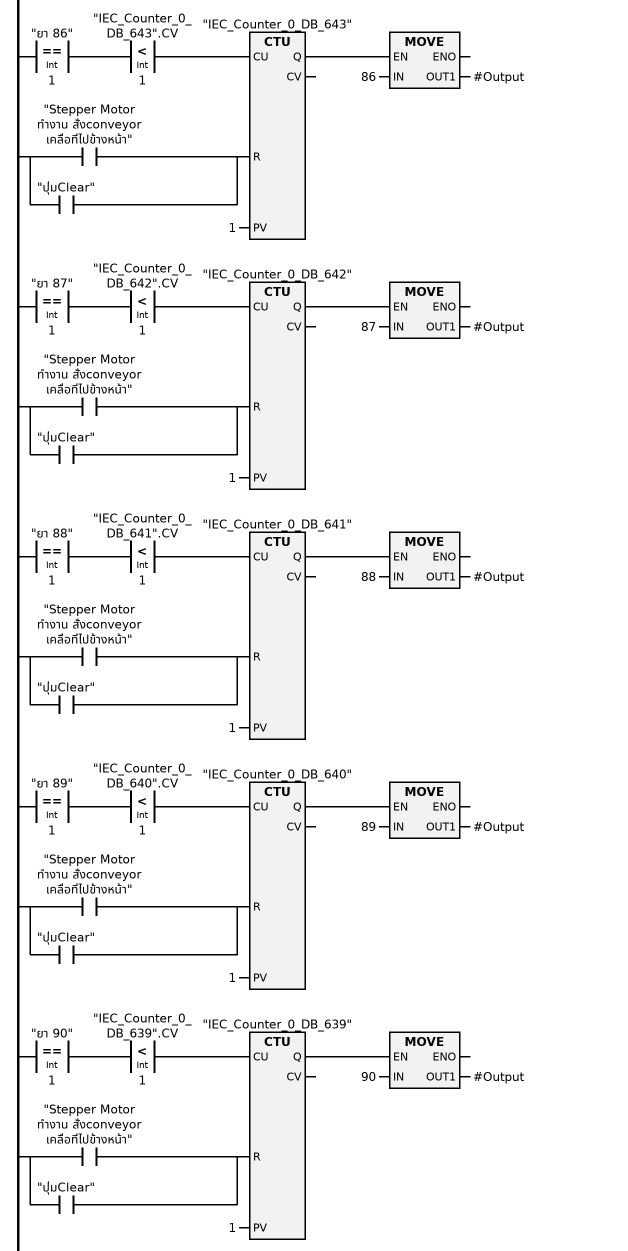
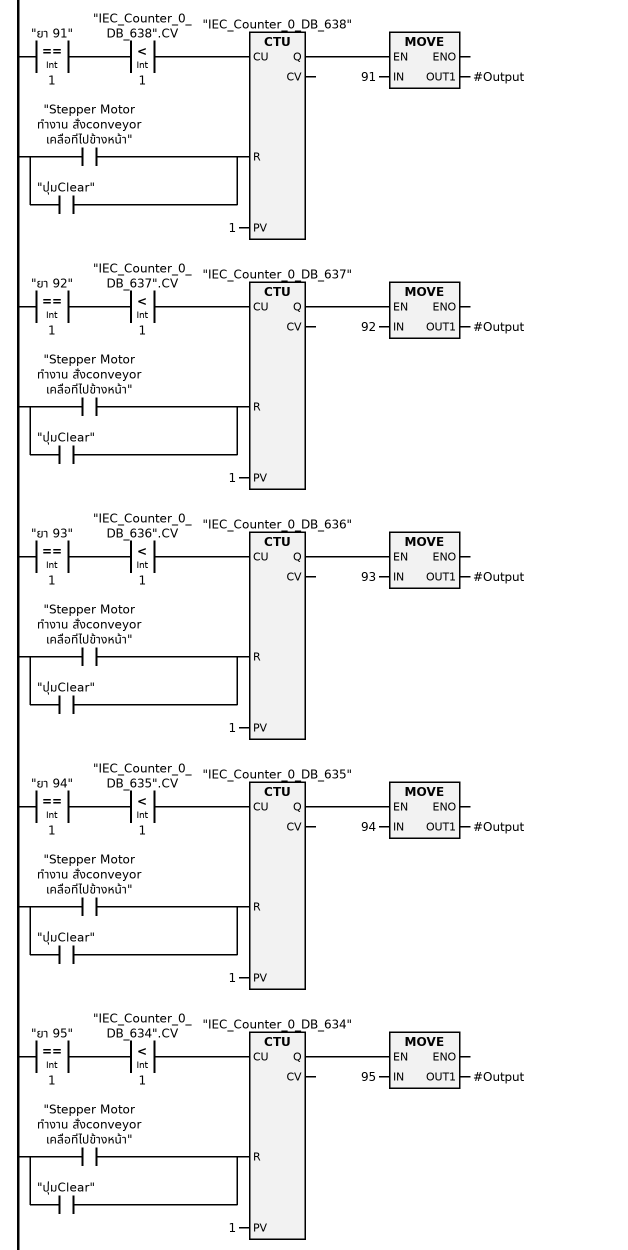
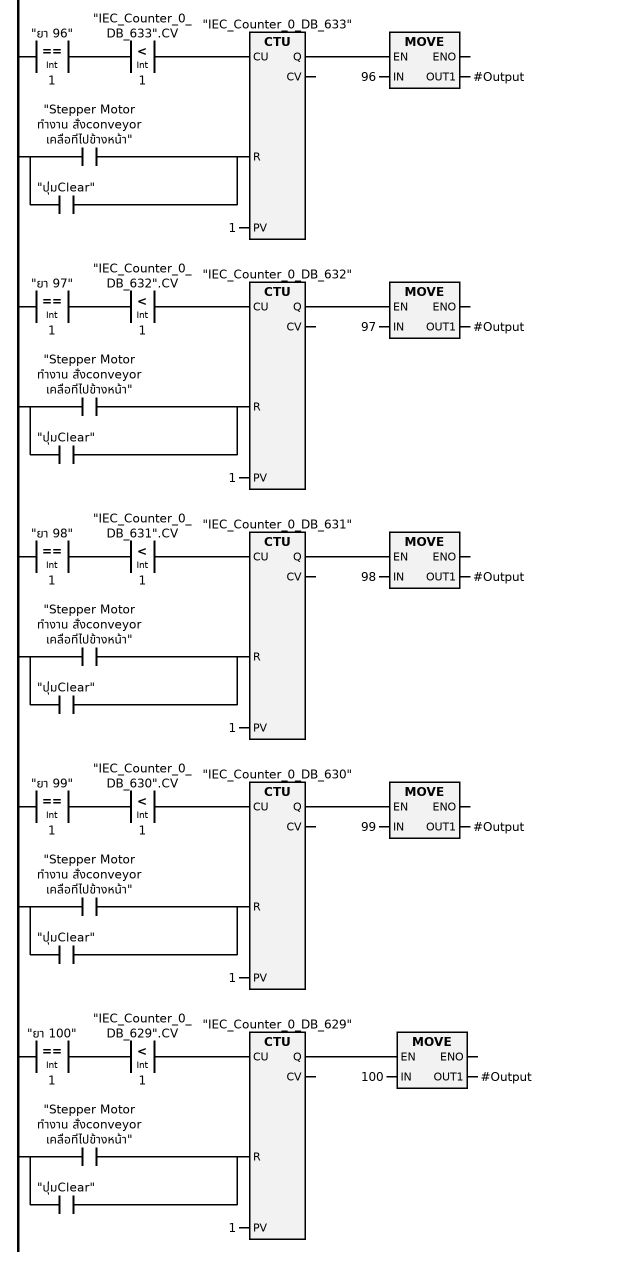
   "IEC_Counter_0_DB_644".CTU(CU := ("ยา 81" = 1) AND ("IEC_Counter_0_DB_644".CV < 1),
                           R := "Stepper Motor ทำงาน สั่งconveyor เคลื่อที่ไปข้างหน้า" OR "ปุ่มClear",
                           PV := 1);
   IF "IEC_Counter_0_DB_644".Q THEN #Output := 81; END_IF;
   "IEC_Counter_0_DB_645".CTU(CU := ("ยา 82" = 1) AND ("IEC_Counter_0_DB_645".CV < 1),
                           R := "Stepper Motor ทำงาน สั่งconveyor เคลื่อที่ไปข้างหน้า" OR "ปุ่มClear",
                           PV := 1);
   IF "IEC_Counter_0_DB_645".Q THEN #Output := 82; END_IF;
   "IEC_Counter_0_DB_647".CTU(CU := ("ยา 83" = 1) AND ("IEC_Counter_0_DB_647".CV < 1),
                           R := "Stepper Motor ทำงาน สั่งconveyor เคลื่อที่ไปข้างหน้า" OR "ปุ่มClear",
                           PV := 1);
   IF "IEC_Counter_0_DB_647".Q THEN #Output := 83; END_IF;
   "IEC_Counter_0_DB_648".CTU(CU := ("ยา 84" = 1) AND ("IEC_Counter_0_DB_648".CV < 1),
                           R := "Stepper Motor ทำงาน สั่งconveyor เคลื่อที่ไปข้างหน้า" OR "ปุ่มClear",
                           PV := 1);
   IF "IEC_Counter_0_DB_648".Q THEN #Output := 84; END_IF;
   "IEC_Counter_0_DB_646".CTU(CU := ("ยา 85" = 1) AND ("IEC_Counter_0_DB_646".CV < 1),
                           R := "Stepper Motor ทำงาน สั่งconveyor เคลื่อที่ไปข้างหน้า" OR "ปุ่มClear",
                           PV := 1);
   IF "IEC_Counter_0_DB_646".Q THEN #Output := 85; END_IF;
   "IEC_Counter_0_DB_643".CTU(CU := ("ยา 86" = 1) AND ("IEC_Counter_0_DB_643".CV < 1),
                           R := "Stepper Motor ทำงาน สั่งconveyor เคลื่อที่ไปข้างหน้า" OR "ปุ่มClear",
                           PV := 1);
   IF "IEC_Counter_0_DB_643".Q THEN #Output := 86; END_IF;
   "IEC_Counter_0_DB_642".CTU(CU := ("ยา 87" = 1) AND ("IEC_Counter_0_DB_642".CV < 1),
                           R := "Stepper Motor ทำงาน สั่งconveyor เคลื่อที่ไปข้างหน้า" OR "ปุ่มClear",
                           PV := 1);
   IF "IEC_Counter_0_DB_642".Q THEN #Output := 87; END_IF;
   "IEC_Counter_0_DB_641".CTU(CU := ("ยา 88" = 1) AND ("IEC_Counter_0_DB_641".CV < 1),
                           R := "Stepper Motor ทำงาน สั่งconveyor เคลื่อที่ไปข้างหน้า" OR "ปุ่มClear",
                           PV := 1);
   IF "IEC_Counter_0_DB_641".Q THEN #Output := 88; END_IF;
   "IEC_Counter_0_DB_640".CTU(CU := ("ยา 89" = 1) AND ("IEC_Counter_0_DB_640".CV < 1),
                           R := "Stepper Motor ทำงาน สั่งconveyor เคลื่อที่ไปข้างหน้า" OR "ปุ่มClear",
                           PV := 1);
   IF "IEC_Counter_0_DB_640".Q THEN #Output := 89; END_IF;
   "IEC_Counter_0_DB_639".CTU(CU := ("ยา 90" = 1) AND ("IEC_Counter_0_DB_639".CV < 1),
                           R := "Stepper Motor ทำงาน สั่งconveyor เคลื่อที่ไปข้างหน้า" OR "ปุ่มClear",
                           PV := 1);
   IF "IEC_Counter_0_DB_639".Q THEN #Output := 90; END_IF;
   "IEC_Counter_0_DB_638".CTU(CU := ("ยา 91" = 1) AND ("IEC_Counter_0_DB_638".CV < 1),
                           R := "Stepper Motor ทำงาน สั่งconveyor เคลื่อที่ไปข้างหน้า" OR "ปุ่มClear",
                           PV := 1);
   IF "IEC_Counter_0_DB_638".Q THEN #Output := 91; END_IF;
   "IEC_Counter_0_DB_637".CTU(CU := ("ยา 92" = 1) AND ("IEC_Counter_0_DB_637".CV < 1),
                           R := "Stepper Motor ทำงาน สั่งconveyor เคลื่อที่ไปข้างหน้า" OR "ปุ่มClear",
                           PV := 1);
   IF "IEC_Counter_0_DB_637".Q THEN #Output := 92; END_IF;
   "IEC_Counter_0_DB_636".CTU(CU := ("ยา 93" = 1) AND ("IEC_Counter_0_DB_636".CV < 1),
                           R := "Stepper Motor ทำงาน สั่งconveyor เคลื่อที่ไปข้างหน้า" OR "ปุ่มClear",
                           PV := 1);
   IF "IEC_Counter_0_DB_636".Q THEN #Output := 93; END_IF;
   "IEC_Counter_0_DB_635".CTU(CU := ("ยา 94" = 1) AND ("IEC_Counter_0_DB_635".CV < 1),
                           R := "Stepper Motor ทำงาน สั่งconveyor เคลื่อที่ไปข้างหน้า" OR "ปุ่มClear",
                           PV := 1);
   IF "IEC_Counter_0_DB_635".Q THEN #Output := 94; END_IF;
   "IEC_Counter_0_DB_634".CTU(CU := ("ยา 95" = 1) AND ("IEC_Counter_0_DB_634".CV < 1),
                           R := "Stepper Motor ทำงาน สั่งconveyor เคลื่อที่ไปข้างหน้า" OR "ปุ่มClear",
                           PV := 1);
   IF "IEC_Counter_0_DB_634".Q THEN #Output := 95; END_IF;
   "IEC_Counter_0_DB_633".CTU(CU := ("ยา 96" = 1) AND ("IEC_Counter_0_DB_633".CV < 1),
                           R := "Stepper Motor ทำงาน สั่งconveyor เคลื่อที่ไปข้างหน้า" OR "ปุ่มClear",
                           PV := 1);
   IF "IEC_Counter_0_DB_633".Q THEN #Output := 96; END_IF;
   "IEC_Counter_0_DB_632".CTU(CU := ("ยา 97" = 1) AND ("IEC_Counter_0_DB_632".CV < 1),
                           R := "Stepper Motor ทำงาน สั่งconveyor เคลื่อที่ไปข้างหน้า" OR "ปุ่มClear",
                           PV := 1);
   IF "IEC_Counter_0_DB_632".Q THEN #Output := 97; END_IF;
   "IEC_Counter_0_DB_631".CTU(CU := ("ยา 98" = 1) AND ("IEC_Counter_0_DB_631".CV < 1),
                           R := "Stepper Motor ทำงาน สั่งconveyor เคลื่อที่ไปข้างหน้า" OR "ปุ่มClear",
                           PV := 1);
   IF "IEC_Counter_0_DB_631".Q THEN #Output := 98; END_IF;
   "IEC_Counter_0_DB_630".CTU(CU := ("ยา 99" = 1) AND ("IEC_Counter_0_DB_630".CV < 1),
                           R := "Stepper Motor ทำงาน สั่งconveyor เคลื่อที่ไปข้างหน้า" OR "ปุ่มClear",
                           PV := 1);
   IF "IEC_Counter_0_DB_630".Q THEN #Output := 99; END_IF;
   "IEC_Counter_0_DB_629".CTU(CU := ("ยา 100" = 1) AND ("IEC_Counter_0_DB_629".CV < 1),
                           R := "Stepper Motor ทำงาน สั่งconveyor เคลื่อที่ไปข้างหน้า" OR "ปุ่มClear",
                           PV := 1);
   IF "IEC_Counter_0_DB_629".Q THEN #Output := 100; END_IF;
END_REGION

REGION Network 6
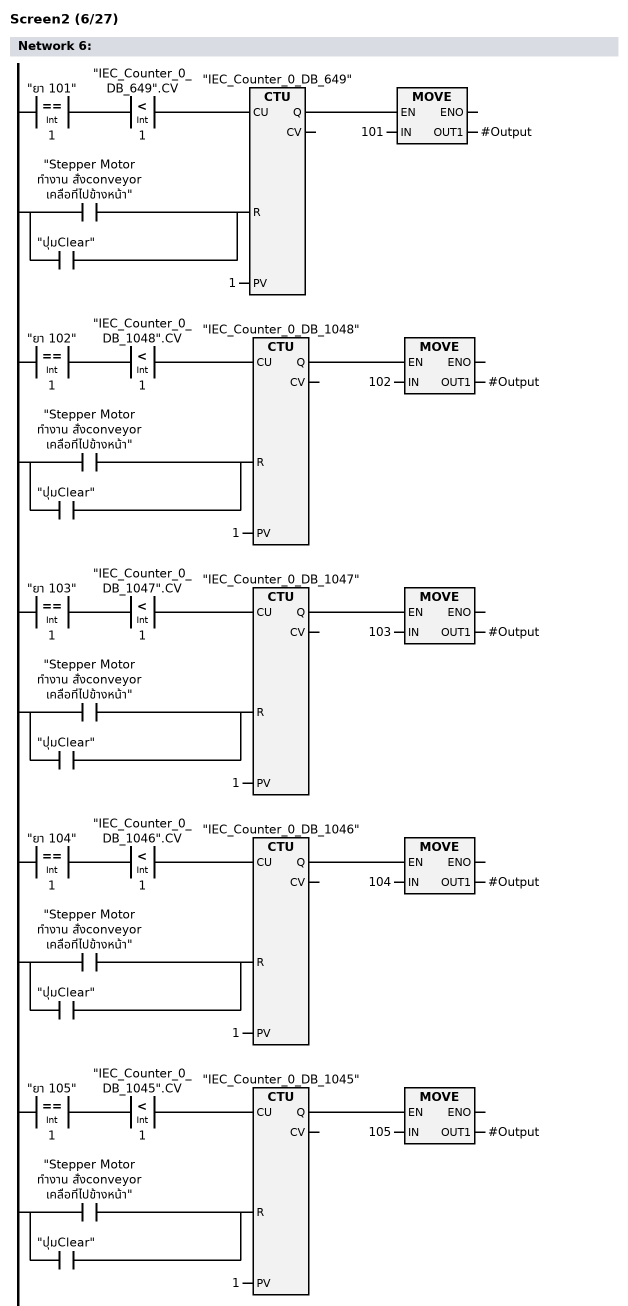
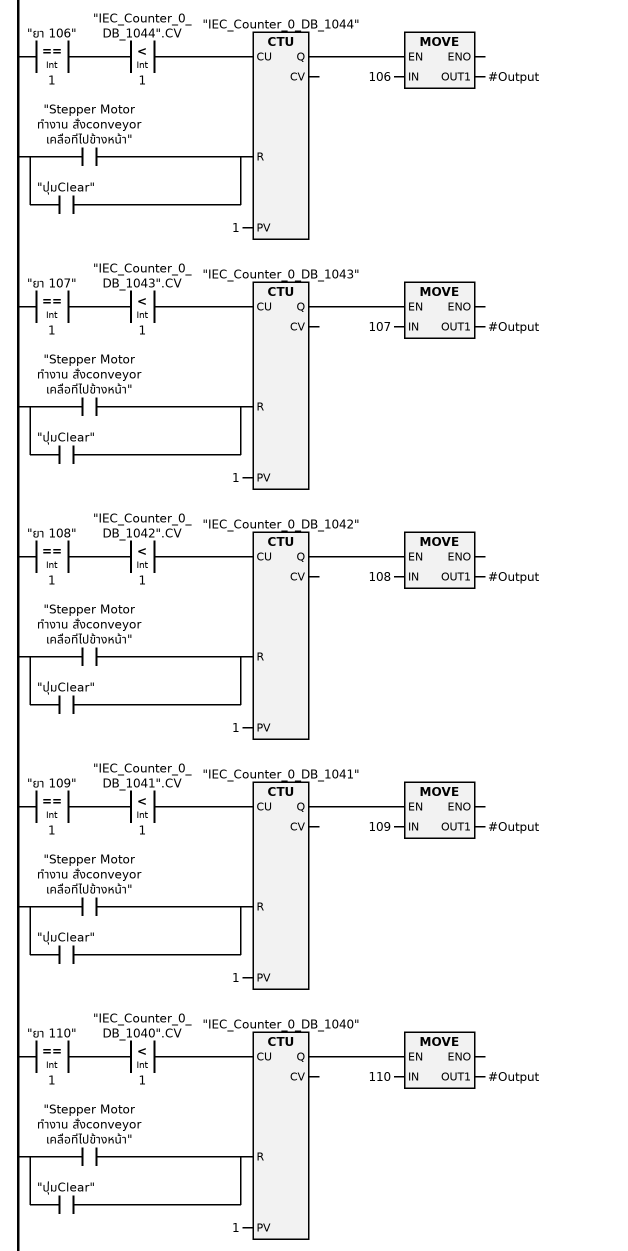
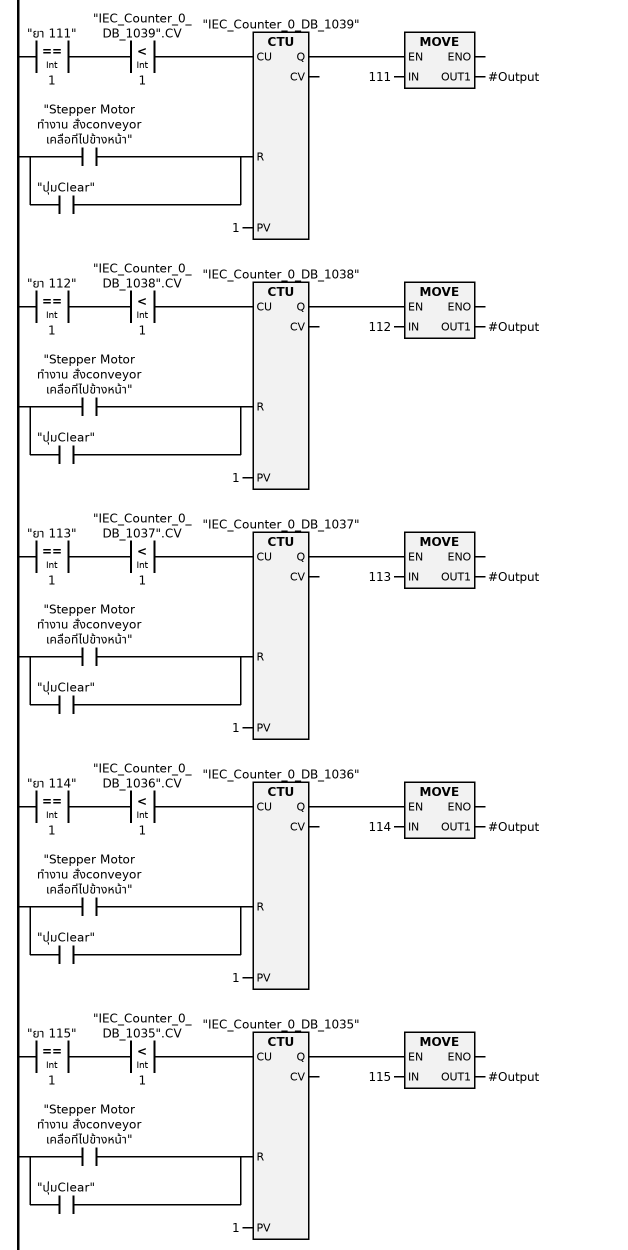
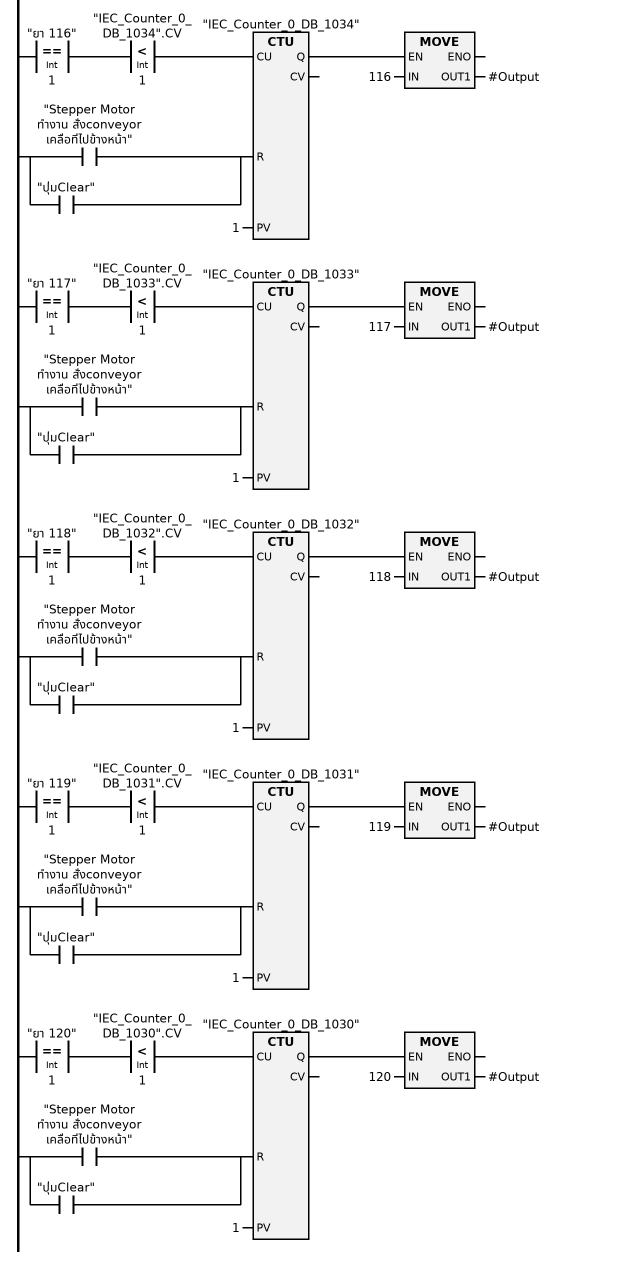
   "IEC_Counter_0_DB_649".CTU(CU := ("ยา 101" = 1) AND ("IEC_Counter_0_DB_649".CV < 1),
                           R := "Stepper Motor ทำงาน สั่งconveyor เคลื่อที่ไปข้างหน้า" OR "ปุ่มClear",
                           PV := 1);
   IF "IEC_Counter_0_DB_649".Q THEN #Output := 101; END_IF;
   "IEC_Counter_0_DB_1048".CTU(CU := ("ยา 102" = 1) AND ("IEC_Counter_0_DB_1048".CV < 1),
                           R := "Stepper Motor ทำงาน สั่งconveyor เคลื่อที่ไปข้างหน้า" OR "ปุ่มClear",
                           PV := 1);
   IF "IEC_Counter_0_DB_1048".Q THEN #Output := 102; END_IF;
   "IEC_Counter_0_DB_1047".CTU(CU := ("ยา 103" = 1) AND ("IEC_Counter_0_DB_1047".CV < 1),
                           R := "Stepper Motor ทำงาน สั่งconveyor เคลื่อที่ไปข้างหน้า" OR "ปุ่มClear",
                           PV := 1);
   IF "IEC_Counter_0_DB_1047".Q THEN #Output := 103; END_IF;
   "IEC_Counter_0_DB_1046".CTU(CU := ("ยา 104" = 1) AND ("IEC_Counter_0_DB_1046".CV < 1),
                           R := "Stepper Motor ทำงาน สั่งconveyor เคลื่อที่ไปข้างหน้า" OR "ปุ่มClear",
                           PV := 1);
   IF "IEC_Counter_0_DB_1046".Q THEN #Output := 104; END_IF;
   "IEC_Counter_0_DB_1045".CTU(CU := ("ยา 105" = 1) AND ("IEC_Counter_0_DB_1045".CV < 1),
                           R := "Stepper Motor ทำงาน สั่งconveyor เคลื่อที่ไปข้างหน้า" OR "ปุ่มClear",
                           PV := 1);
   IF "IEC_Counter_0_DB_1045".Q THEN #Output := 105; END_IF;
   "IEC_Counter_0_DB_1044".CTU(CU := ("ยา 106" = 1) AND ("IEC_Counter_0_DB_1044".CV < 1),
                           R := "Stepper Motor ทำงาน สั่งconveyor เคลื่อที่ไปข้างหน้า" OR "ปุ่มClear",
                           PV := 1);
   IF "IEC_Counter_0_DB_1044".Q THEN #Output := 106; END_IF;
   "IEC_Counter_0_DB_1043".CTU(CU := ("ยา 107" = 1) AND ("IEC_Counter_0_DB_1043".CV < 1),
                           R := "Stepper Motor ทำงาน สั่งconveyor เคลื่อที่ไปข้างหน้า" OR "ปุ่มClear",
                           PV := 1);
   IF "IEC_Counter_0_DB_1043".Q THEN #Output := 107; END_IF;
   "IEC_Counter_0_DB_1042".CTU(CU := ("ยา 108" = 1) AND ("IEC_Counter_0_DB_1042".CV < 1),
                           R := "Stepper Motor ทำงาน สั่งconveyor เคลื่อที่ไปข้างหน้า" OR "ปุ่มClear",
                           PV := 1);
   IF "IEC_Counter_0_DB_1042".Q THEN #Output := 108; END_IF;
   "IEC_Counter_0_DB_1041".CTU(CU := ("ยา 109" = 1) AND ("IEC_Counter_0_DB_1041".CV < 1),
                           R := "Stepper Motor ทำงาน สั่งconveyor เคลื่อที่ไปข้างหน้า" OR "ปุ่มClear",
                           PV := 1);
   IF "IEC_Counter_0_DB_1041".Q THEN #Output := 109; END_IF;
   "IEC_Counter_0_DB_1040".CTU(CU := ("ยา 110" = 1) AND ("IEC_Counter_0_DB_1040".CV < 1),
                           R := "Stepper Motor ทำงาน สั่งconveyor เคลื่อที่ไปข้างหน้า" OR "ปุ่มClear",
                           PV := 1);
   IF "IEC_Counter_0_DB_1040".Q THEN #Output := 110; END_IF;
   "IEC_Counter_0_DB_1039".CTU(CU := ("ยา 111" = 1) AND ("IEC_Counter_0_DB_1039".CV < 1),
                           R := "Stepper Motor ทำงาน สั่งconveyor เคลื่อที่ไปข้างหน้า" OR "ปุ่มClear",
                           PV := 1);
   IF "IEC_Counter_0_DB_1039".Q THEN #Output := 111; END_IF;
   "IEC_Counter_0_DB_1038".CTU(CU := ("ยา 112" = 1) AND ("IEC_Counter_0_DB_1038".CV < 1),
                           R := "Stepper Motor ทำงาน สั่งconveyor เคลื่อที่ไปข้างหน้า" OR "ปุ่มClear",
                           PV := 1);
   IF "IEC_Counter_0_DB_1038".Q THEN #Output := 112; END_IF;
   "IEC_Counter_0_DB_1037".CTU(CU := ("ยา 113" = 1) AND ("IEC_Counter_0_DB_1037".CV < 1),
                           R := "Stepper Motor ทำงาน สั่งconveyor เคลื่อที่ไปข้างหน้า" OR "ปุ่มClear",
                           PV := 1);
   IF "IEC_Counter_0_DB_1037".Q THEN #Output := 113; END_IF;
   "IEC_Counter_0_DB_1036".CTU(CU := ("ยา 114" = 1) AND ("IEC_Counter_0_DB_1036".CV < 1),
                           R := "Stepper Motor ทำงาน สั่งconveyor เคลื่อที่ไปข้างหน้า" OR "ปุ่มClear",
                           PV := 1);
   IF "IEC_Counter_0_DB_1036".Q THEN #Output := 114; END_IF;
   "IEC_Counter_0_DB_1035".CTU(CU := ("ยา 115" = 1) AND ("IEC_Counter_0_DB_1035".CV < 1),
                           R := "Stepper Motor ทำงาน สั่งconveyor เคลื่อที่ไปข้างหน้า" OR "ปุ่มClear",
                           PV := 1);
   IF "IEC_Counter_0_DB_1035".Q THEN #Output := 115; END_IF;
   "IEC_Counter_0_DB_1034".CTU(CU := ("ยา 116" = 1) AND ("IEC_Counter_0_DB_1034".CV < 1),
                           R := "Stepper Motor ทำงาน สั่งconveyor เคลื่อที่ไปข้างหน้า" OR "ปุ่มClear",
                           PV := 1);
   IF "IEC_Counter_0_DB_1034".Q THEN #Output := 116; END_IF;
   "IEC_Counter_0_DB_1033".CTU(CU := ("ยา 117" = 1) AND ("IEC_Counter_0_DB_1033".CV < 1),
                           R := "Stepper Motor ทำงาน สั่งconveyor เคลื่อที่ไปข้างหน้า" OR "ปุ่มClear",
                           PV := 1);
   IF "IEC_Counter_0_DB_1033".Q THEN #Output := 117; END_IF;
   "IEC_Counter_0_DB_1032".CTU(CU := ("ยา 118" = 1) AND ("IEC_Counter_0_DB_1032".CV < 1),
                           R := "Stepper Motor ทำงาน สั่งconveyor เคลื่อที่ไปข้างหน้า" OR "ปุ่มClear",
                           PV := 1);
   IF "IEC_Counter_0_DB_1032".Q THEN #Output := 118; END_IF;
   "IEC_Counter_0_DB_1031".CTU(CU := ("ยา 119" = 1) AND ("IEC_Counter_0_DB_1031".CV < 1),
                           R := "Stepper Motor ทำงาน สั่งconveyor เคลื่อที่ไปข้างหน้า" OR "ปุ่มClear",
                           PV := 1);
   IF "IEC_Counter_0_DB_1031".Q THEN #Output := 119; END_IF;
   "IEC_Counter_0_DB_1030".CTU(CU := ("ยา 120" = 1) AND ("IEC_Counter_0_DB_1030".CV < 1),
                           R := "Stepper Motor ทำงาน สั่งconveyor เคลื่อที่ไปข้างหน้า" OR "ปุ่มClear",
                           PV := 1);
   IF "IEC_Counter_0_DB_1030".Q THEN #Output := 120; END_IF;
END_REGION

REGION Network 7
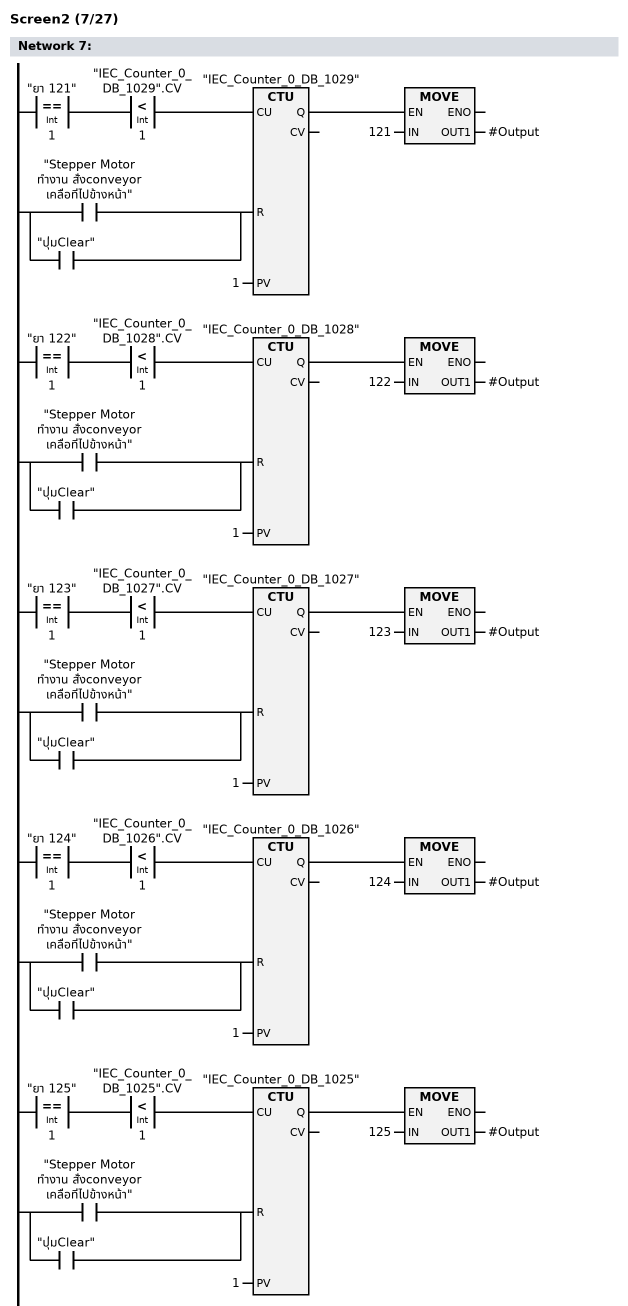
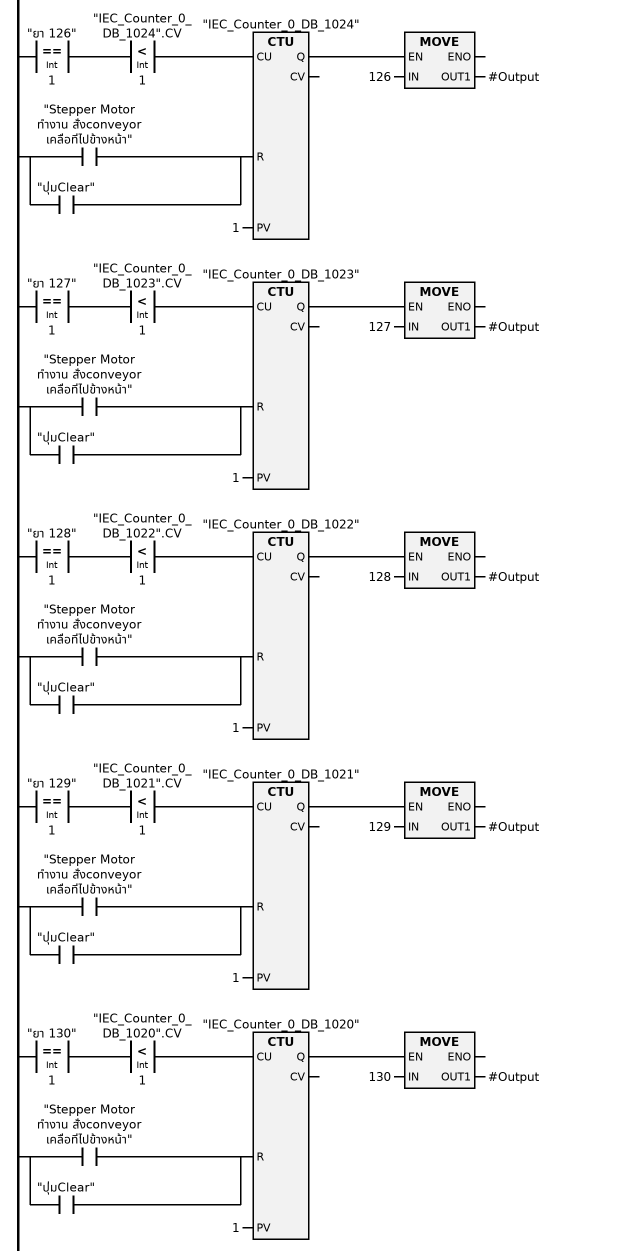
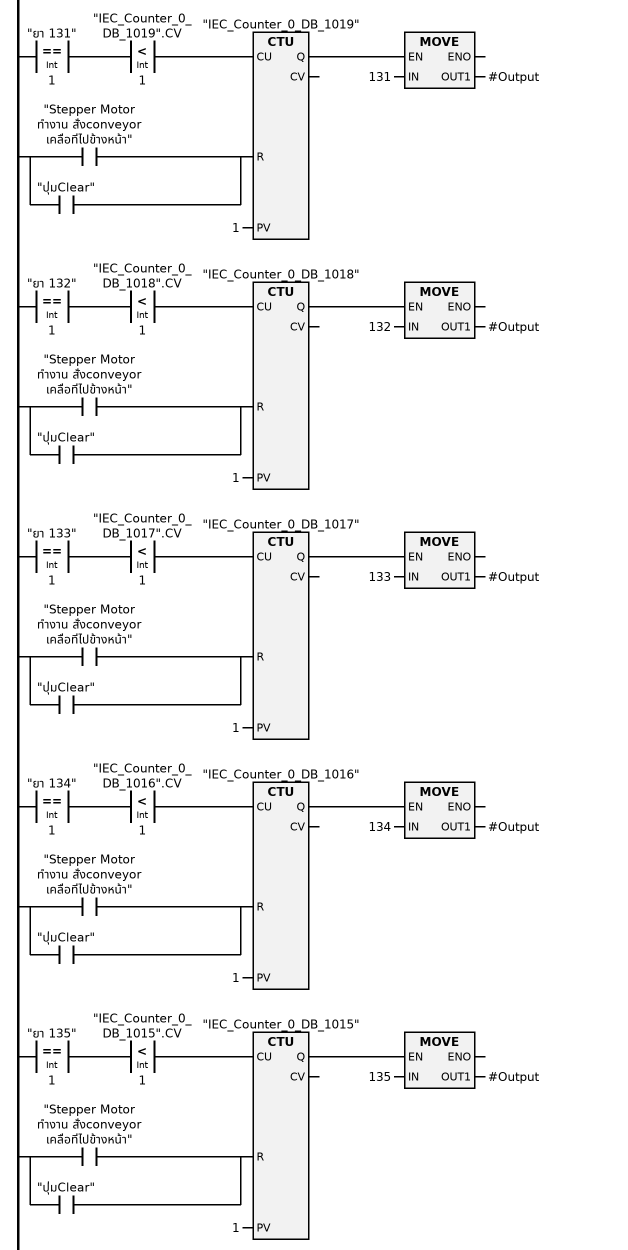
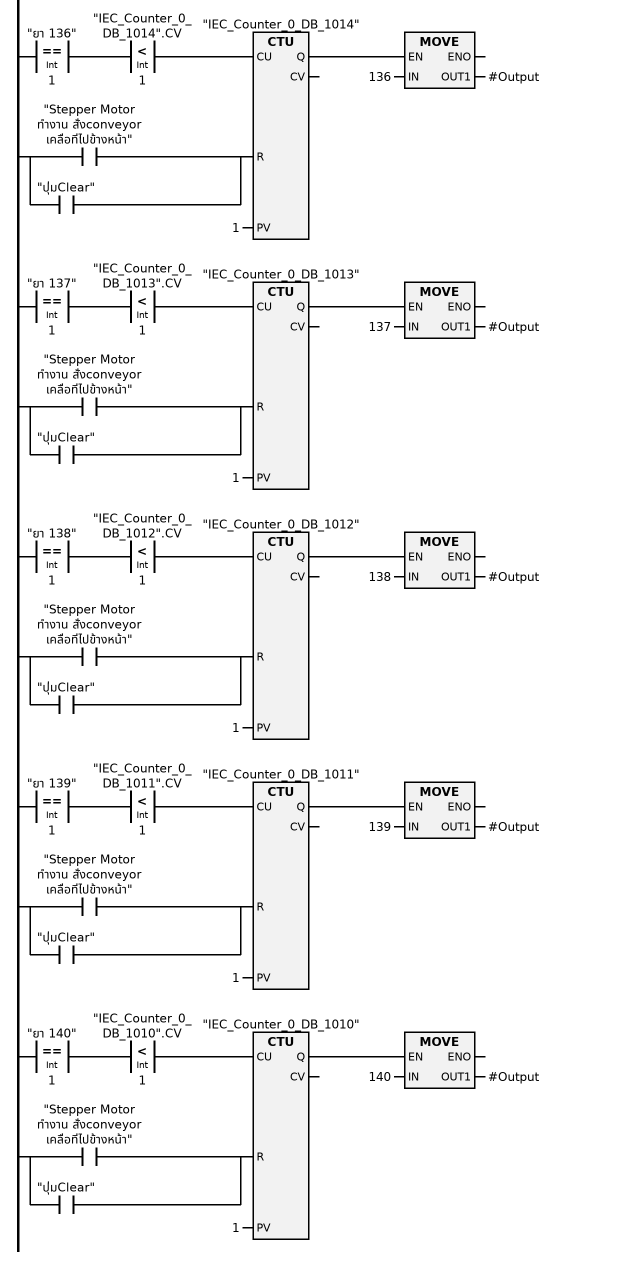
   "IEC_Counter_0_DB_1029".CTU(CU := ("ยา 121" = 1) AND ("IEC_Counter_0_DB_1029".CV < 1),
                           R := "Stepper Motor ทำงาน สั่งconveyor เคลื่อที่ไปข้างหน้า" OR "ปุ่มClear",
                           PV := 1);
   IF "IEC_Counter_0_DB_1029".Q THEN #Output := 121; END_IF;
   "IEC_Counter_0_DB_1028".CTU(CU := ("ยา 122" = 1) AND ("IEC_Counter_0_DB_1028".CV < 1),
                           R := "Stepper Motor ทำงาน สั่งconveyor เคลื่อที่ไปข้างหน้า" OR "ปุ่มClear",
                           PV := 1);
   IF "IEC_Counter_0_DB_1028".Q THEN #Output := 122; END_IF;
   "IEC_Counter_0_DB_1027".CTU(CU := ("ยา 123" = 1) AND ("IEC_Counter_0_DB_1027".CV < 1),
                           R := "Stepper Motor ทำงาน สั่งconveyor เคลื่อที่ไปข้างหน้า" OR "ปุ่มClear",
                           PV := 1);
   IF "IEC_Counter_0_DB_1027".Q THEN #Output := 123; END_IF;
   "IEC_Counter_0_DB_1026".CTU(CU := ("ยา 124" = 1) AND ("IEC_Counter_0_DB_1026".CV < 1),
                           R := "Stepper Motor ทำงาน สั่งconveyor เคลื่อที่ไปข้างหน้า" OR "ปุ่มClear",
                           PV := 1);
   IF "IEC_Counter_0_DB_1026".Q THEN #Output := 124; END_IF;
   "IEC_Counter_0_DB_1025".CTU(CU := ("ยา 125" = 1) AND ("IEC_Counter_0_DB_1025".CV < 1),
                           R := "Stepper Motor ทำงาน สั่งconveyor เคลื่อที่ไปข้างหน้า" OR "ปุ่มClear",
                           PV := 1);
   IF "IEC_Counter_0_DB_1025".Q THEN #Output := 125; END_IF;
   "IEC_Counter_0_DB_1024".CTU(CU := ("ยา 126" = 1) AND ("IEC_Counter_0_DB_1024".CV < 1),
                           R := "Stepper Motor ทำงาน สั่งconveyor เคลื่อที่ไปข้างหน้า" OR "ปุ่มClear",
                           PV := 1);
   IF "IEC_Counter_0_DB_1024".Q THEN #Output := 126; END_IF;
   "IEC_Counter_0_DB_1023".CTU(CU := ("ยา 127" = 1) AND ("IEC_Counter_0_DB_1023".CV < 1),
                           R := "Stepper Motor ทำงาน สั่งconveyor เคลื่อที่ไปข้างหน้า" OR "ปุ่มClear",
                           PV := 1);
   IF "IEC_Counter_0_DB_1023".Q THEN #Output := 127; END_IF;
   "IEC_Counter_0_DB_1022".CTU(CU := ("ยา 128" = 1) AND ("IEC_Counter_0_DB_1022".CV < 1),
                           R := "Stepper Motor ทำงาน สั่งconveyor เคลื่อที่ไปข้างหน้า" OR "ปุ่มClear",
                           PV := 1);
   IF "IEC_Counter_0_DB_1022".Q THEN #Output := 128; END_IF;
   "IEC_Counter_0_DB_1021".CTU(CU := ("ยา 129" = 1) AND ("IEC_Counter_0_DB_1021".CV < 1),
                           R := "Stepper Motor ทำงาน สั่งconveyor เคลื่อที่ไปข้างหน้า" OR "ปุ่มClear",
                           PV := 1);
   IF "IEC_Counter_0_DB_1021".Q THEN #Output := 129; END_IF;
   "IEC_Counter_0_DB_1020".CTU(CU := ("ยา 130" = 1) AND ("IEC_Counter_0_DB_1020".CV < 1),
                           R := "Stepper Motor ทำงาน สั่งconveyor เคลื่อที่ไปข้างหน้า" OR "ปุ่มClear",
                           PV := 1);
   IF "IEC_Counter_0_DB_1020".Q THEN #Output := 130; END_IF;
   "IEC_Counter_0_DB_1019".CTU(CU := ("ยา 131" = 1) AND ("IEC_Counter_0_DB_1019".CV < 1),
                           R := "Stepper Motor ทำงาน สั่งconveyor เคลื่อที่ไปข้างหน้า" OR "ปุ่มClear",
                           PV := 1);
   IF "IEC_Counter_0_DB_1019".Q THEN #Output := 131; END_IF;
   "IEC_Counter_0_DB_1018".CTU(CU := ("ยา 132" = 1) AND ("IEC_Counter_0_DB_1018".CV < 1),
                           R := "Stepper Motor ทำงาน สั่งconveyor เคลื่อที่ไปข้างหน้า" OR "ปุ่มClear",
                           PV := 1);
   IF "IEC_Counter_0_DB_1018".Q THEN #Output := 132; END_IF;
   "IEC_Counter_0_DB_1017".CTU(CU := ("ยา 133" = 1) AND ("IEC_Counter_0_DB_1017".CV < 1),
                           R := "Stepper Motor ทำงาน สั่งconveyor เคลื่อที่ไปข้างหน้า" OR "ปุ่มClear",
                           PV := 1);
   IF "IEC_Counter_0_DB_1017".Q THEN #Output := 133; END_IF;
   "IEC_Counter_0_DB_1016".CTU(CU := ("ยา 134" = 1) AND ("IEC_Counter_0_DB_1016".CV < 1),
                           R := "Stepper Motor ทำงาน สั่งconveyor เคลื่อที่ไปข้างหน้า" OR "ปุ่มClear",
                           PV := 1);
   IF "IEC_Counter_0_DB_1016".Q THEN #Output := 134; END_IF;
   "IEC_Counter_0_DB_1015".CTU(CU := ("ยา 135" = 1) AND ("IEC_Counter_0_DB_1015".CV < 1),
                           R := "Stepper Motor ทำงาน สั่งconveyor เคลื่อที่ไปข้างหน้า" OR "ปุ่มClear",
                           PV := 1);
   IF "IEC_Counter_0_DB_1015".Q THEN #Output := 135; END_IF;
   "IEC_Counter_0_DB_1014".CTU(CU := ("ยา 136" = 1) AND ("IEC_Counter_0_DB_1014".CV < 1),
                           R := "Stepper Motor ทำงาน สั่งconveyor เคลื่อที่ไปข้างหน้า" OR "ปุ่มClear",
                           PV := 1);
   IF "IEC_Counter_0_DB_1014".Q THEN #Output := 136; END_IF;
   "IEC_Counter_0_DB_1013".CTU(CU := ("ยา 137" = 1) AND ("IEC_Counter_0_DB_1013".CV < 1),
                           R := "Stepper Motor ทำงาน สั่งconveyor เคลื่อที่ไปข้างหน้า" OR "ปุ่มClear",
                           PV := 1);
   IF "IEC_Counter_0_DB_1013".Q THEN #Output := 137; END_IF;
   "IEC_Counter_0_DB_1012".CTU(CU := ("ยา 138" = 1) AND ("IEC_Counter_0_DB_1012".CV < 1),
                           R := "Stepper Motor ทำงาน สั่งconveyor เคลื่อที่ไปข้างหน้า" OR "ปุ่มClear",
                           PV := 1);
   IF "IEC_Counter_0_DB_1012".Q THEN #Output := 138; END_IF;
   "IEC_Counter_0_DB_1011".CTU(CU := ("ยา 139" = 1) AND ("IEC_Counter_0_DB_1011".CV < 1),
                           R := "Stepper Motor ทำงาน สั่งconveyor เคลื่อที่ไปข้างหน้า" OR "ปุ่มClear",
                           PV := 1);
   IF "IEC_Counter_0_DB_1011".Q THEN #Output := 139; END_IF;
   "IEC_Counter_0_DB_1010".CTU(CU := ("ยา 140" = 1) AND ("IEC_Counter_0_DB_1010".CV < 1),
                           R := "Stepper Motor ทำงาน สั่งconveyor เคลื่อที่ไปข้างหน้า" OR "ปุ่มClear",
                           PV := 1);
   IF "IEC_Counter_0_DB_1010".Q THEN #Output := 140; END_IF;
END_REGION

REGION Network 8
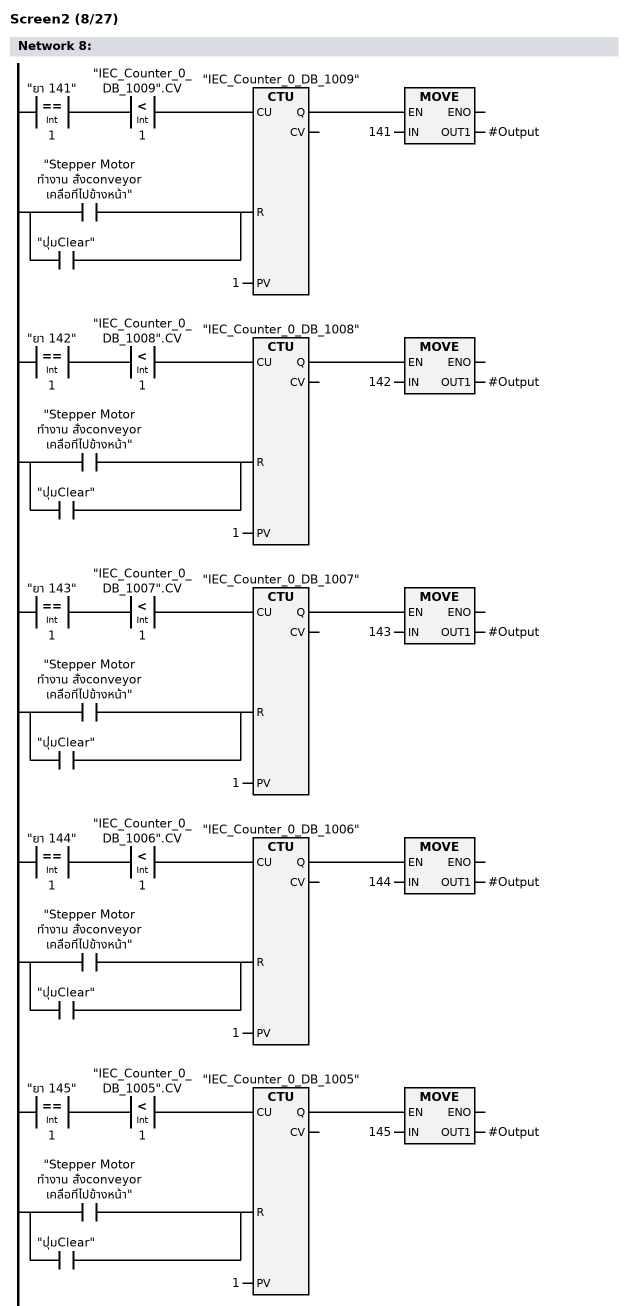
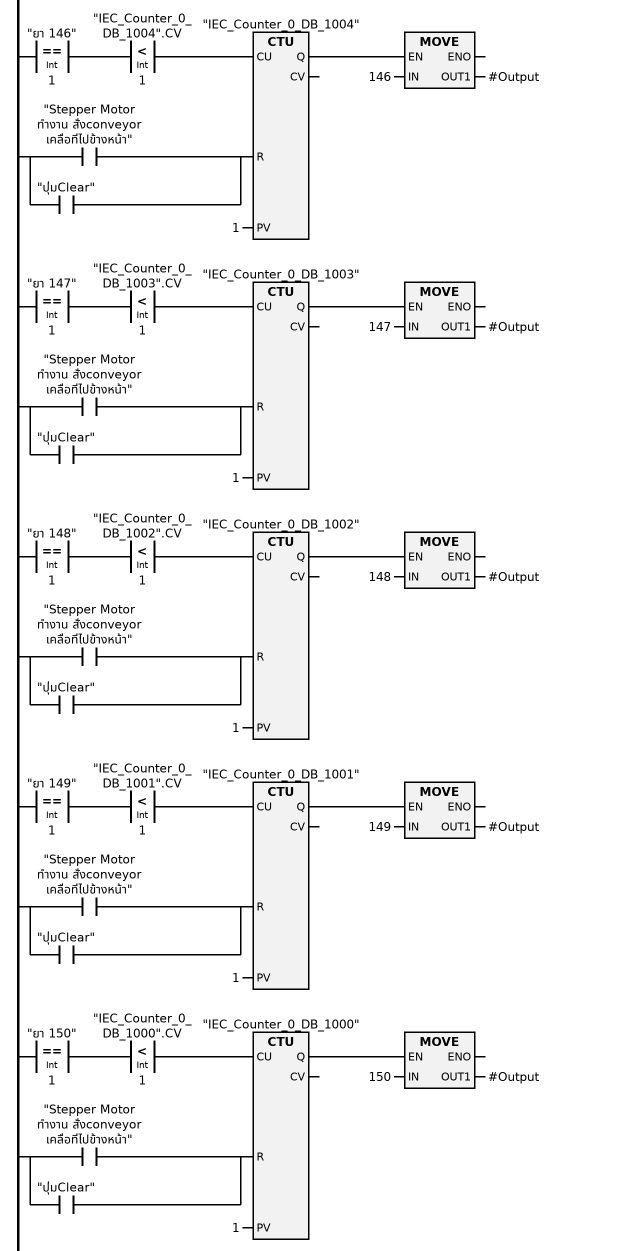
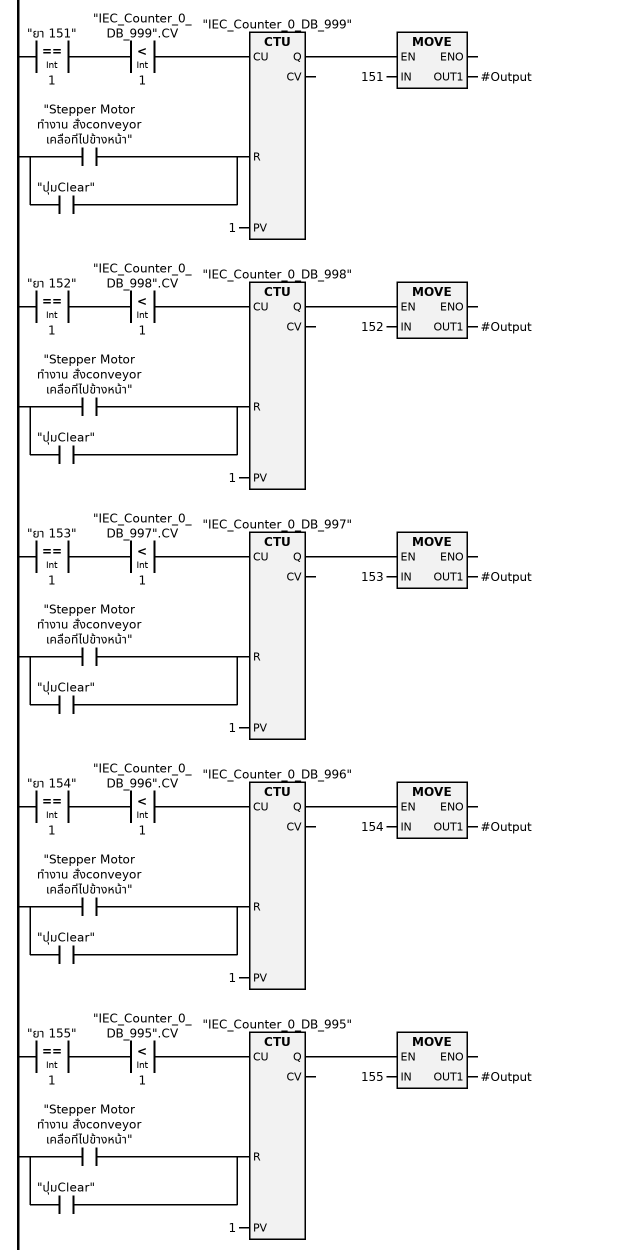
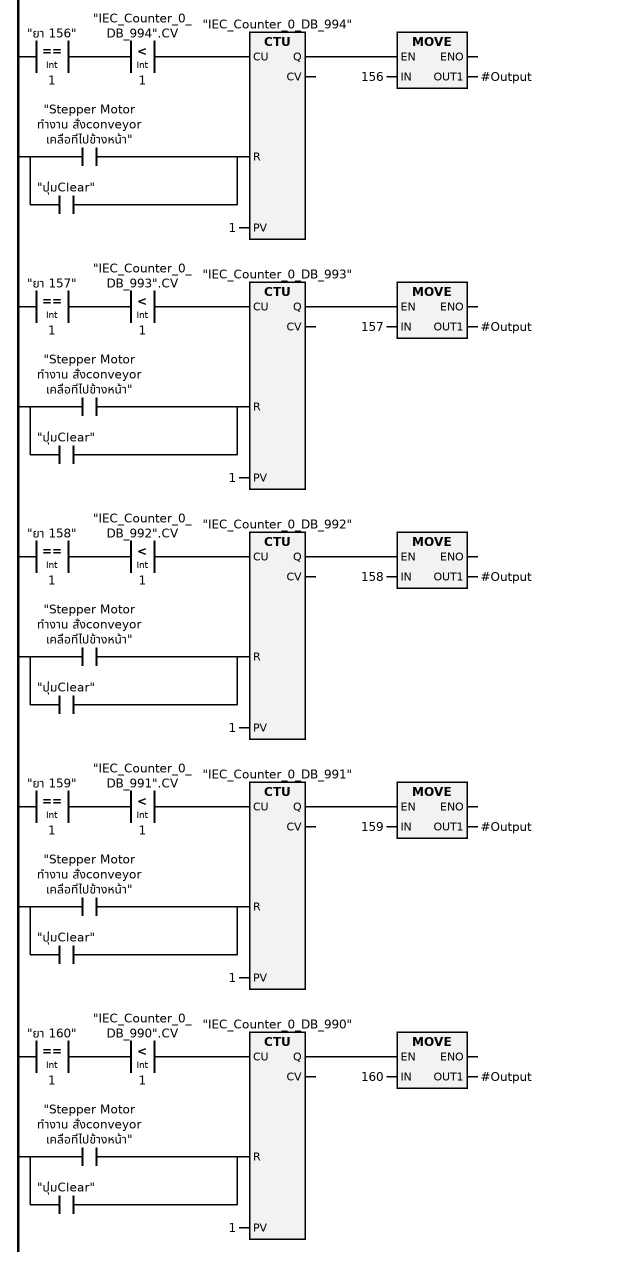
   "IEC_Counter_0_DB_1009".CTU(CU := ("ยา 141" = 1) AND ("IEC_Counter_0_DB_1009".CV < 1),
                           R := "Stepper Motor ทำงาน สั่งconveyor เคลื่อที่ไปข้างหน้า" OR "ปุ่มClear",
                           PV := 1);
   IF "IEC_Counter_0_DB_1009".Q THEN #Output := 141; END_IF;
   "IEC_Counter_0_DB_1008".CTU(CU := ("ยา 142" = 1) AND ("IEC_Counter_0_DB_1008".CV < 1),
                           R := "Stepper Motor ทำงาน สั่งconveyor เคลื่อที่ไปข้างหน้า" OR "ปุ่มClear",
                           PV := 1);
   IF "IEC_Counter_0_DB_1008".Q THEN #Output := 142; END_IF;
   "IEC_Counter_0_DB_1007".CTU(CU := ("ยา 143" = 1) AND ("IEC_Counter_0_DB_1007".CV < 1),
                           R := "Stepper Motor ทำงาน สั่งconveyor เคลื่อที่ไปข้างหน้า" OR "ปุ่มClear",
                           PV := 1);
   IF "IEC_Counter_0_DB_1007".Q THEN #Output := 143; END_IF;
   "IEC_Counter_0_DB_1006".CTU(CU := ("ยา 144" = 1) AND ("IEC_Counter_0_DB_1006".CV < 1),
                           R := "Stepper Motor ทำงาน สั่งconveyor เคลื่อที่ไปข้างหน้า" OR "ปุ่มClear",
                           PV := 1);
   IF "IEC_Counter_0_DB_1006".Q THEN #Output := 144; END_IF;
   "IEC_Counter_0_DB_1005".CTU(CU := ("ยา 145" = 1) AND ("IEC_Counter_0_DB_1005".CV < 1),
                           R := "Stepper Motor ทำงาน สั่งconveyor เคลื่อที่ไปข้างหน้า" OR "ปุ่มClear",
                           PV := 1);
   IF "IEC_Counter_0_DB_1005".Q THEN #Output := 145; END_IF;
   "IEC_Counter_0_DB_1004".CTU(CU := ("ยา 146" = 1) AND ("IEC_Counter_0_DB_1004".CV < 1),
                           R := "Stepper Motor ทำงาน สั่งconveyor เคลื่อที่ไปข้างหน้า" OR "ปุ่มClear",
                           PV := 1);
   IF "IEC_Counter_0_DB_1004".Q THEN #Output := 146; END_IF;
   "IEC_Counter_0_DB_1003".CTU(CU := ("ยา 147" = 1) AND ("IEC_Counter_0_DB_1003".CV < 1),
                           R := "Stepper Motor ทำงาน สั่งconveyor เคลื่อที่ไปข้างหน้า" OR "ปุ่มClear",
                           PV := 1);
   IF "IEC_Counter_0_DB_1003".Q THEN #Output := 147; END_IF;
   "IEC_Counter_0_DB_1002".CTU(CU := ("ยา 148" = 1) AND ("IEC_Counter_0_DB_1002".CV < 1),
                           R := "Stepper Motor ทำงาน สั่งconveyor เคลื่อที่ไปข้างหน้า" OR "ปุ่มClear",
                           PV := 1);
   IF "IEC_Counter_0_DB_1002".Q THEN #Output := 148; END_IF;
   "IEC_Counter_0_DB_1001".CTU(CU := ("ยา 149" = 1) AND ("IEC_Counter_0_DB_1001".CV < 1),
                           R := "Stepper Motor ทำงาน สั่งconveyor เคลื่อที่ไปข้างหน้า" OR "ปุ่มClear",
                           PV := 1);
   IF "IEC_Counter_0_DB_1001".Q THEN #Output := 149; END_IF;
   "IEC_Counter_0_DB_1000".CTU(CU := ("ยา 150" = 1) AND ("IEC_Counter_0_DB_1000".CV < 1),
                           R := "Stepper Motor ทำงาน สั่งconveyor เคลื่อที่ไปข้างหน้า" OR "ปุ่มClear",
                           PV := 1);
   IF "IEC_Counter_0_DB_1000".Q THEN #Output := 150; END_IF;
   "IEC_Counter_0_DB_999".CTU(CU := ("ยา 151" = 1) AND ("IEC_Counter_0_DB_999".CV < 1),
                           R := "Stepper Motor ทำงาน สั่งconveyor เคลื่อที่ไปข้างหน้า" OR "ปุ่มClear",
                           PV := 1);
   IF "IEC_Counter_0_DB_999".Q THEN #Output := 151; END_IF;
   "IEC_Counter_0_DB_998".CTU(CU := ("ยา 152" = 1) AND ("IEC_Counter_0_DB_998".CV < 1),
                           R := "Stepper Motor ทำงาน สั่งconveyor เคลื่อที่ไปข้างหน้า" OR "ปุ่มClear",
                           PV := 1);
   IF "IEC_Counter_0_DB_998".Q THEN #Output := 152; END_IF;
   "IEC_Counter_0_DB_997".CTU(CU := ("ยา 153" = 1) AND ("IEC_Counter_0_DB_997".CV < 1),
                           R := "Stepper Motor ทำงาน สั่งconveyor เคลื่อที่ไปข้างหน้า" OR "ปุ่มClear",
                           PV := 1);
   IF "IEC_Counter_0_DB_997".Q THEN #Output := 153; END_IF;
   "IEC_Counter_0_DB_996".CTU(CU := ("ยา 154" = 1) AND ("IEC_Counter_0_DB_996".CV < 1),
                           R := "Stepper Motor ทำงาน สั่งconveyor เคลื่อที่ไปข้างหน้า" OR "ปุ่มClear",
                           PV := 1);
   IF "IEC_Counter_0_DB_996".Q THEN #Output := 154; END_IF;
   "IEC_Counter_0_DB_995".CTU(CU := ("ยา 155" = 1) AND ("IEC_Counter_0_DB_995".CV < 1),
                           R := "Stepper Motor ทำงาน สั่งconveyor เคลื่อที่ไปข้างหน้า" OR "ปุ่มClear",
                           PV := 1);
   IF "IEC_Counter_0_DB_995".Q THEN #Output := 155; END_IF;
   "IEC_Counter_0_DB_994".CTU(CU := ("ยา 156" = 1) AND ("IEC_Counter_0_DB_994".CV < 1),
                           R := "Stepper Motor ทำงาน สั่งconveyor เคลื่อที่ไปข้างหน้า" OR "ปุ่มClear",
                           PV := 1);
   IF "IEC_Counter_0_DB_994".Q THEN #Output := 156; END_IF;
   "IEC_Counter_0_DB_993".CTU(CU := ("ยา 157" = 1) AND ("IEC_Counter_0_DB_993".CV < 1),
                           R := "Stepper Motor ทำงาน สั่งconveyor เคลื่อที่ไปข้างหน้า" OR "ปุ่มClear",
                           PV := 1);
   IF "IEC_Counter_0_DB_993".Q THEN #Output := 157; END_IF;
   "IEC_Counter_0_DB_992".CTU(CU := ("ยา 158" = 1) AND ("IEC_Counter_0_DB_992".CV < 1),
                           R := "Stepper Motor ทำงาน สั่งconveyor เคลื่อที่ไปข้างหน้า" OR "ปุ่มClear",
                           PV := 1);
   IF "IEC_Counter_0_DB_992".Q THEN #Output := 158; END_IF;
   "IEC_Counter_0_DB_991".CTU(CU := ("ยา 159" = 1) AND ("IEC_Counter_0_DB_991".CV < 1),
                           R := "Stepper Motor ทำงาน สั่งconveyor เคลื่อที่ไปข้างหน้า" OR "ปุ่มClear",
                           PV := 1);
   IF "IEC_Counter_0_DB_991".Q THEN #Output := 159; END_IF;
   "IEC_Counter_0_DB_990".CTU(CU := ("ยา 160" = 1) AND ("IEC_Counter_0_DB_990".CV < 1),
                           R := "Stepper Motor ทำงาน สั่งconveyor เคลื่อที่ไปข้างหน้า" OR "ปุ่มClear",
                           PV := 1);
   IF "IEC_Counter_0_DB_990".Q THEN #Output := 160; END_IF;
END_REGION

REGION Network 9
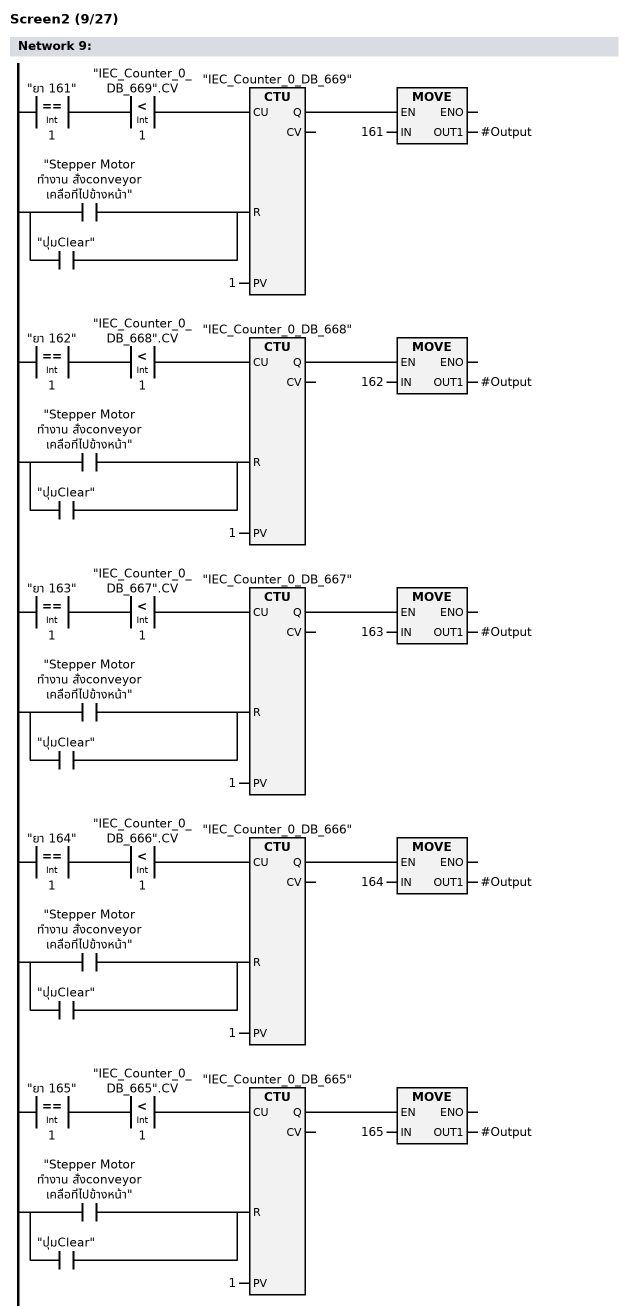
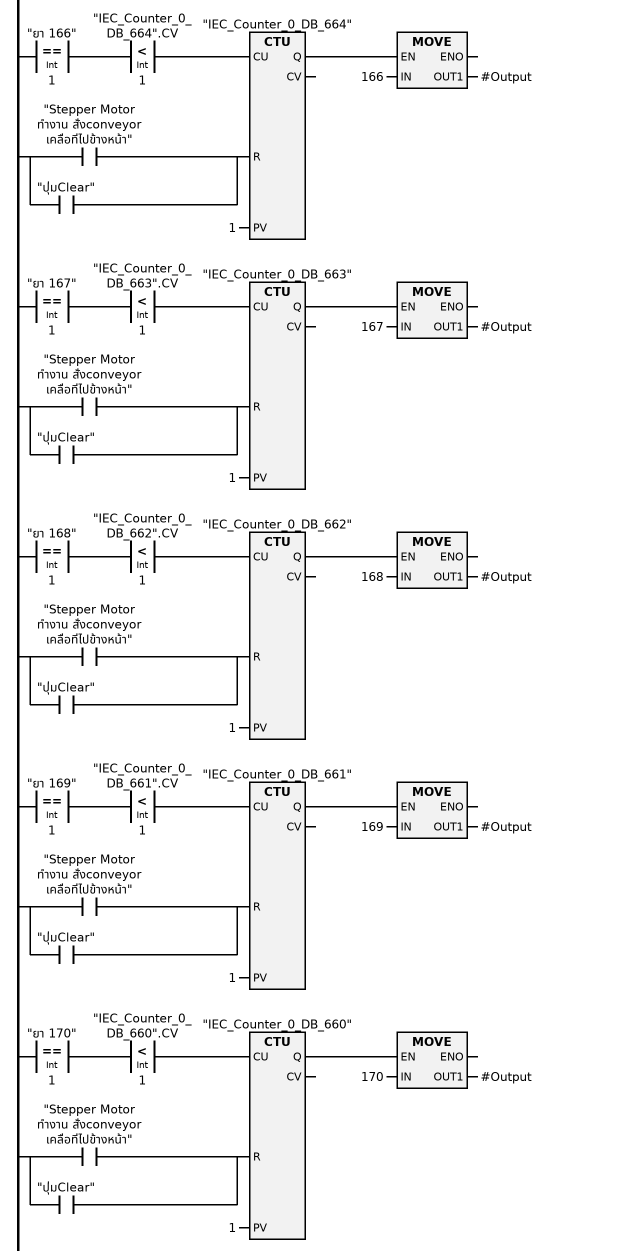
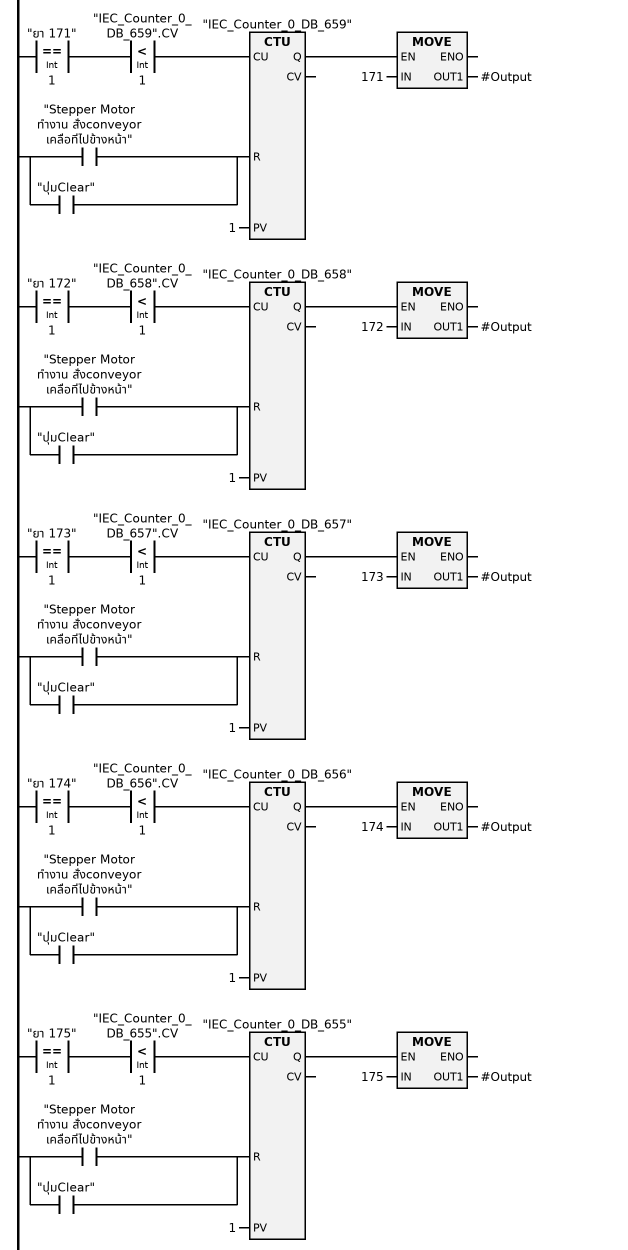
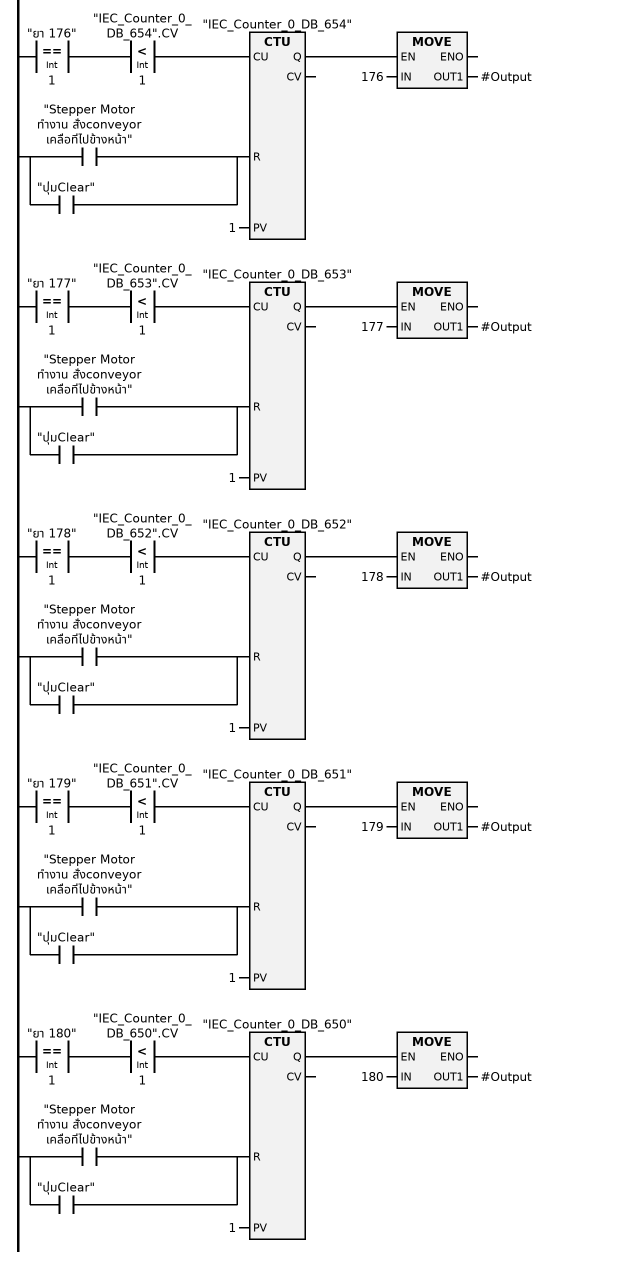
   "IEC_Counter_0_DB_669".CTU(CU := ("ยา 161" = 1) AND ("IEC_Counter_0_DB_669".CV < 1),
                           R := "Stepper Motor ทำงาน สั่งconveyor เคลื่อที่ไปข้างหน้า" OR "ปุ่มClear",
                           PV := 1);
   IF "IEC_Counter_0_DB_669".Q THEN #Output := 161; END_IF;
   "IEC_Counter_0_DB_668".CTU(CU := ("ยา 162" = 1) AND ("IEC_Counter_0_DB_668".CV < 1),
                           R := "Stepper Motor ทำงาน สั่งconveyor เคลื่อที่ไปข้างหน้า" OR "ปุ่มClear",
                           PV := 1);
   IF "IEC_Counter_0_DB_668".Q THEN #Output := 162; END_IF;
   "IEC_Counter_0_DB_667".CTU(CU := ("ยา 163" = 1) AND ("IEC_Counter_0_DB_667".CV < 1),
                           R := "Stepper Motor ทำงาน สั่งconveyor เคลื่อที่ไปข้างหน้า" OR "ปุ่มClear",
                           PV := 1);
   IF "IEC_Counter_0_DB_667".Q THEN #Output := 163; END_IF;
   "IEC_Counter_0_DB_666".CTU(CU := ("ยา 164" = 1) AND ("IEC_Counter_0_DB_666".CV < 1),
                           R := "Stepper Motor ทำงาน สั่งconveyor เคลื่อที่ไปข้างหน้า" OR "ปุ่มClear",
                           PV := 1);
   IF "IEC_Counter_0_DB_666".Q THEN #Output := 164; END_IF;
   "IEC_Counter_0_DB_665".CTU(CU := ("ยา 165" = 1) AND ("IEC_Counter_0_DB_665".CV < 1),
                           R := "Stepper Motor ทำงาน สั่งconveyor เคลื่อที่ไปข้างหน้า" OR "ปุ่มClear",
                           PV := 1);
   IF "IEC_Counter_0_DB_665".Q THEN #Output := 165; END_IF;
   "IEC_Counter_0_DB_664".CTU(CU := ("ยา 166" = 1) AND ("IEC_Counter_0_DB_664".CV < 1),
                           R := "Stepper Motor ทำงาน สั่งconveyor เคลื่อที่ไปข้างหน้า" OR "ปุ่มClear",
                           PV := 1);
   IF "IEC_Counter_0_DB_664".Q THEN #Output := 166; END_IF;
   "IEC_Counter_0_DB_663".CTU(CU := ("ยา 167" = 1) AND ("IEC_Counter_0_DB_663".CV < 1),
                           R := "Stepper Motor ทำงาน สั่งconveyor เคลื่อที่ไปข้างหน้า" OR "ปุ่มClear",
                           PV := 1);
   IF "IEC_Counter_0_DB_663".Q THEN #Output := 167; END_IF;
   "IEC_Counter_0_DB_662".CTU(CU := ("ยา 168" = 1) AND ("IEC_Counter_0_DB_662".CV < 1),
                           R := "Stepper Motor ทำงาน สั่งconveyor เคลื่อที่ไปข้างหน้า" OR "ปุ่มClear",
                           PV := 1);
   IF "IEC_Counter_0_DB_662".Q THEN #Output := 168; END_IF;
   "IEC_Counter_0_DB_661".CTU(CU := ("ยา 169" = 1) AND ("IEC_Counter_0_DB_661".CV < 1),
                           R := "Stepper Motor ทำงาน สั่งconveyor เคลื่อที่ไปข้างหน้า" OR "ปุ่มClear",
                           PV := 1);
   IF "IEC_Counter_0_DB_661".Q THEN #Output := 169; END_IF;
   "IEC_Counter_0_DB_660".CTU(CU := ("ยา 170" = 1) AND ("IEC_Counter_0_DB_660".CV < 1),
                           R := "Stepper Motor ทำงาน สั่งconveyor เคลื่อที่ไปข้างหน้า" OR "ปุ่มClear",
                           PV := 1);
   IF "IEC_Counter_0_DB_660".Q THEN #Output := 170; END_IF;
   "IEC_Counter_0_DB_659".CTU(CU := ("ยา 171" = 1) AND ("IEC_Counter_0_DB_659".CV < 1),
                           R := "Stepper Motor ทำงาน สั่งconveyor เคลื่อที่ไปข้างหน้า" OR "ปุ่มClear",
                           PV := 1);
   IF "IEC_Counter_0_DB_659".Q THEN #Output := 171; END_IF;
   "IEC_Counter_0_DB_658".CTU(CU := ("ยา 172" = 1) AND ("IEC_Counter_0_DB_658".CV < 1),
                           R := "Stepper Motor ทำงาน สั่งconveyor เคลื่อที่ไปข้างหน้า" OR "ปุ่มClear",
                           PV := 1);
   IF "IEC_Counter_0_DB_658".Q THEN #Output := 172; END_IF;
   "IEC_Counter_0_DB_657".CTU(CU := ("ยา 173" = 1) AND ("IEC_Counter_0_DB_657".CV < 1),
                           R := "Stepper Motor ทำงาน สั่งconveyor เคลื่อที่ไปข้างหน้า" OR "ปุ่มClear",
                           PV := 1);
   IF "IEC_Counter_0_DB_657".Q THEN #Output := 173; END_IF;
   "IEC_Counter_0_DB_656".CTU(CU := ("ยา 174" = 1) AND ("IEC_Counter_0_DB_656".CV < 1),
                           R := "Stepper Motor ทำงาน สั่งconveyor เคลื่อที่ไปข้างหน้า" OR "ปุ่มClear",
                           PV := 1);
   IF "IEC_Counter_0_DB_656".Q THEN #Output := 174; END_IF;
   "IEC_Counter_0_DB_655".CTU(CU := ("ยา 175" = 1) AND ("IEC_Counter_0_DB_655".CV < 1),
                           R := "Stepper Motor ทำงาน สั่งconveyor เคลื่อที่ไปข้างหน้า" OR "ปุ่มClear",
                           PV := 1);
   IF "IEC_Counter_0_DB_655".Q THEN #Output := 175; END_IF;
   "IEC_Counter_0_DB_654".CTU(CU := ("ยา 176" = 1) AND ("IEC_Counter_0_DB_654".CV < 1),
                           R := "Stepper Motor ทำงาน สั่งconveyor เคลื่อที่ไปข้างหน้า" OR "ปุ่มClear",
                           PV := 1);
   IF "IEC_Counter_0_DB_654".Q THEN #Output := 176; END_IF;
   "IEC_Counter_0_DB_653".CTU(CU := ("ยา 177" = 1) AND ("IEC_Counter_0_DB_653".CV < 1),
                           R := "Stepper Motor ทำงาน สั่งconveyor เคลื่อที่ไปข้างหน้า" OR "ปุ่มClear",
                           PV := 1);
   IF "IEC_Counter_0_DB_653".Q THEN #Output := 177; END_IF;
   "IEC_Counter_0_DB_652".CTU(CU := ("ยา 178" = 1) AND ("IEC_Counter_0_DB_652".CV < 1),
                           R := "Stepper Motor ทำงาน สั่งconveyor เคลื่อที่ไปข้างหน้า" OR "ปุ่มClear",
                           PV := 1);
   IF "IEC_Counter_0_DB_652".Q THEN #Output := 178; END_IF;
   "IEC_Counter_0_DB_651".CTU(CU := ("ยา 179" = 1) AND ("IEC_Counter_0_DB_651".CV < 1),
                           R := "Stepper Motor ทำงาน สั่งconveyor เคลื่อที่ไปข้างหน้า" OR "ปุ่มClear",
                           PV := 1);
   IF "IEC_Counter_0_DB_651".Q THEN #Output := 179; END_IF;
   "IEC_Counter_0_DB_650".CTU(CU := ("ยา 180" = 1) AND ("IEC_Counter_0_DB_650".CV < 1),
                           R := "Stepper Motor ทำงาน สั่งconveyor เคลื่อที่ไปข้างหน้า" OR "ปุ่มClear",
                           PV := 1);
   IF "IEC_Counter_0_DB_650".Q THEN #Output := 180; END_IF;
END_REGION

REGION Network 10
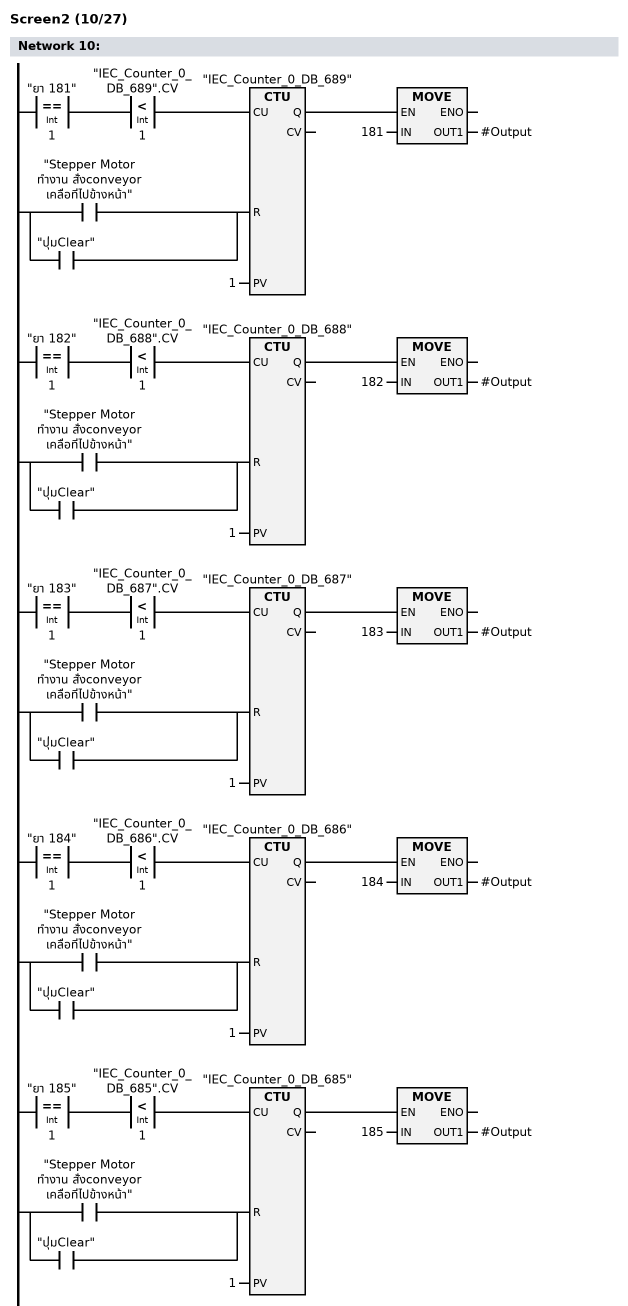
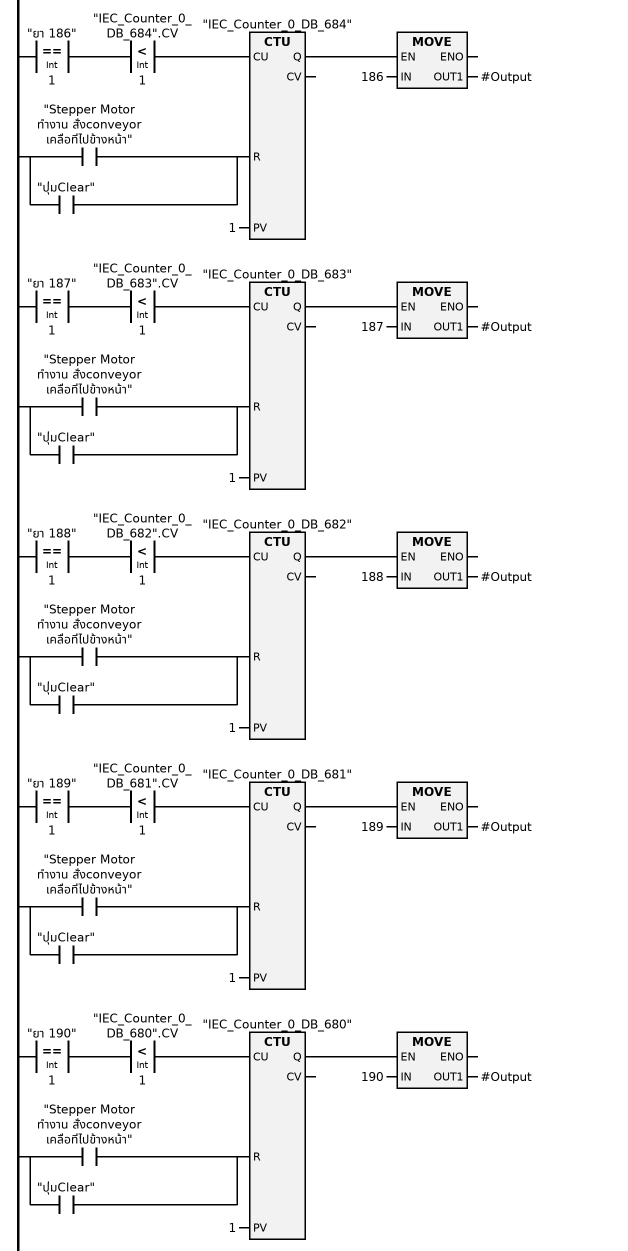
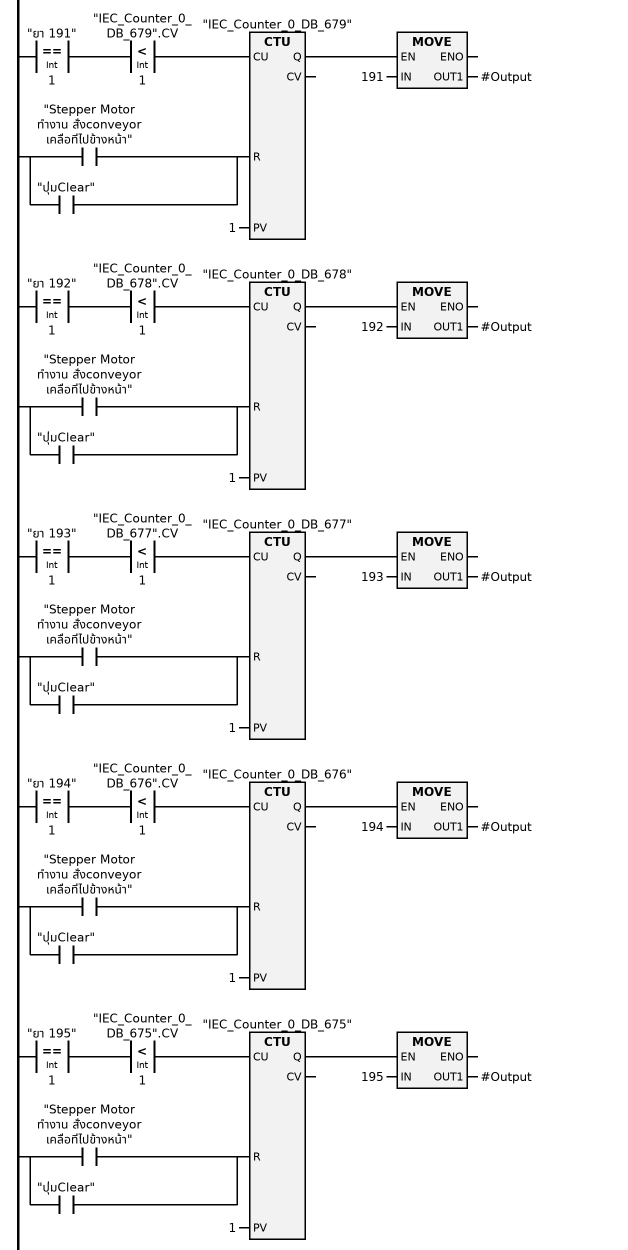
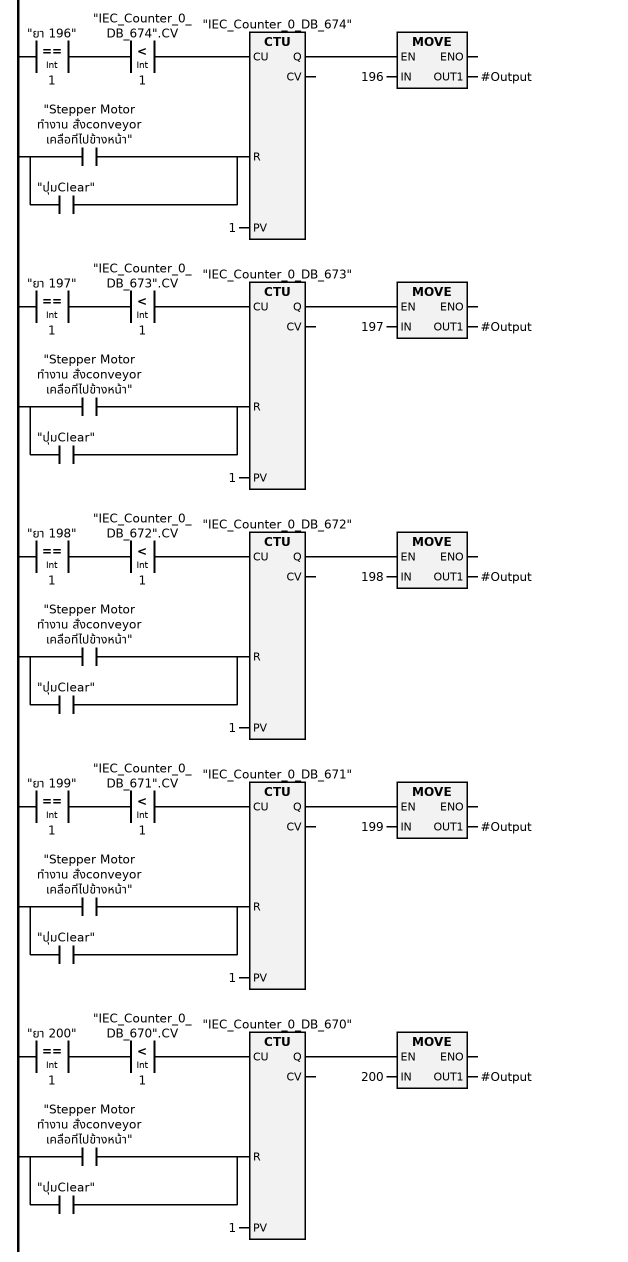
   "IEC_Counter_0_DB_689".CTU(CU := ("ยา 181" = 1) AND ("IEC_Counter_0_DB_689".CV < 1),
                           R := "Stepper Motor ทำงาน สั่งconveyor เคลื่อที่ไปข้างหน้า" OR "ปุ่มClear",
                           PV := 1);
   IF "IEC_Counter_0_DB_689".Q THEN #Output := 181; END_IF;
   "IEC_Counter_0_DB_688".CTU(CU := ("ยา 182" = 1) AND ("IEC_Counter_0_DB_688".CV < 1),
                           R := "Stepper Motor ทำงาน สั่งconveyor เคลื่อที่ไปข้างหน้า" OR "ปุ่มClear",
                           PV := 1);
   IF "IEC_Counter_0_DB_688".Q THEN #Output := 182; END_IF;
   "IEC_Counter_0_DB_687".CTU(CU := ("ยา 183" = 1) AND ("IEC_Counter_0_DB_687".CV < 1),
                           R := "Stepper Motor ทำงาน สั่งconveyor เคลื่อที่ไปข้างหน้า" OR "ปุ่มClear",
                           PV := 1);
   IF "IEC_Counter_0_DB_687".Q THEN #Output := 183; END_IF;
   "IEC_Counter_0_DB_686".CTU(CU := ("ยา 184" = 1) AND ("IEC_Counter_0_DB_686".CV < 1),
                           R := "Stepper Motor ทำงาน สั่งconveyor เคลื่อที่ไปข้างหน้า" OR "ปุ่มClear",
                           PV := 1);
   IF "IEC_Counter_0_DB_686".Q THEN #Output := 184; END_IF;
   "IEC_Counter_0_DB_685".CTU(CU := ("ยา 185" = 1) AND ("IEC_Counter_0_DB_685".CV < 1),
                           R := "Stepper Motor ทำงาน สั่งconveyor เคลื่อที่ไปข้างหน้า" OR "ปุ่มClear",
                           PV := 1);
   IF "IEC_Counter_0_DB_685".Q THEN #Output := 185; END_IF;
   "IEC_Counter_0_DB_684".CTU(CU := ("ยา 186" = 1) AND ("IEC_Counter_0_DB_684".CV < 1),
                           R := "Stepper Motor ทำงาน สั่งconveyor เคลื่อที่ไปข้างหน้า" OR "ปุ่มClear",
                           PV := 1);
   IF "IEC_Counter_0_DB_684".Q THEN #Output := 186; END_IF;
   "IEC_Counter_0_DB_683".CTU(CU := ("ยา 187" = 1) AND ("IEC_Counter_0_DB_683".CV < 1),
                           R := "Stepper Motor ทำงาน สั่งconveyor เคลื่อที่ไปข้างหน้า" OR "ปุ่มClear",
                           PV := 1);
   IF "IEC_Counter_0_DB_683".Q THEN #Output := 187; END_IF;
   "IEC_Counter_0_DB_682".CTU(CU := ("ยา 188" = 1) AND ("IEC_Counter_0_DB_682".CV < 1),
                           R := "Stepper Motor ทำงาน สั่งconveyor เคลื่อที่ไปข้างหน้า" OR "ปุ่มClear",
                           PV := 1);
   IF "IEC_Counter_0_DB_682".Q THEN #Output := 188; END_IF;
   "IEC_Counter_0_DB_681".CTU(CU := ("ยา 189" = 1) AND ("IEC_Counter_0_DB_681".CV < 1),
                           R := "Stepper Motor ทำงาน สั่งconveyor เคลื่อที่ไปข้างหน้า" OR "ปุ่มClear",
                           PV := 1);
   IF "IEC_Counter_0_DB_681".Q THEN #Output := 189; END_IF;
   "IEC_Counter_0_DB_680".CTU(CU := ("ยา 190" = 1) AND ("IEC_Counter_0_DB_680".CV < 1),
                           R := "Stepper Motor ทำงาน สั่งconveyor เคลื่อที่ไปข้างหน้า" OR "ปุ่มClear",
                           PV := 1);
   IF "IEC_Counter_0_DB_680".Q THEN #Output := 190; END_IF;
   "IEC_Counter_0_DB_679".CTU(CU := ("ยา 191" = 1) AND ("IEC_Counter_0_DB_679".CV < 1),
                           R := "Stepper Motor ทำงาน สั่งconveyor เคลื่อที่ไปข้างหน้า" OR "ปุ่มClear",
                           PV := 1);
   IF "IEC_Counter_0_DB_679".Q THEN #Output := 191; END_IF;
   "IEC_Counter_0_DB_678".CTU(CU := ("ยา 192" = 1) AND ("IEC_Counter_0_DB_678".CV < 1),
                           R := "Stepper Motor ทำงาน สั่งconveyor เคลื่อที่ไปข้างหน้า" OR "ปุ่มClear",
                           PV := 1);
   IF "IEC_Counter_0_DB_678".Q THEN #Output := 192; END_IF;
   "IEC_Counter_0_DB_677".CTU(CU := ("ยา 193" = 1) AND ("IEC_Counter_0_DB_677".CV < 1),
                           R := "Stepper Motor ทำงาน สั่งconveyor เคลื่อที่ไปข้างหน้า" OR "ปุ่มClear",
                           PV := 1);
   IF "IEC_Counter_0_DB_677".Q THEN #Output := 193; END_IF;
   "IEC_Counter_0_DB_676".CTU(CU := ("ยา 194" = 1) AND ("IEC_Counter_0_DB_676".CV < 1),
                           R := "Stepper Motor ทำงาน สั่งconveyor เคลื่อที่ไปข้างหน้า" OR "ปุ่มClear",
                           PV := 1);
   IF "IEC_Counter_0_DB_676".Q THEN #Output := 194; END_IF;
   "IEC_Counter_0_DB_675".CTU(CU := ("ยา 195" = 1) AND ("IEC_Counter_0_DB_675".CV < 1),
                           R := "Stepper Motor ทำงาน สั่งconveyor เคลื่อที่ไปข้างหน้า" OR "ปุ่มClear",
                           PV := 1);
   IF "IEC_Counter_0_DB_675".Q THEN #Output := 195; END_IF;
   "IEC_Counter_0_DB_674".CTU(CU := ("ยา 196" = 1) AND ("IEC_Counter_0_DB_674".CV < 1),
                           R := "Stepper Motor ทำงาน สั่งconveyor เคลื่อที่ไปข้างหน้า" OR "ปุ่มClear",
                           PV := 1);
   IF "IEC_Counter_0_DB_674".Q THEN #Output := 196; END_IF;
   "IEC_Counter_0_DB_673".CTU(CU := ("ยา 197" = 1) AND ("IEC_Counter_0_DB_673".CV < 1),
                           R := "Stepper Motor ทำงาน สั่งconveyor เคลื่อที่ไปข้างหน้า" OR "ปุ่มClear",
                           PV := 1);
   IF "IEC_Counter_0_DB_673".Q THEN #Output := 197; END_IF;
   "IEC_Counter_0_DB_672".CTU(CU := ("ยา 198" = 1) AND ("IEC_Counter_0_DB_672".CV < 1),
                           R := "Stepper Motor ทำงาน สั่งconveyor เคลื่อที่ไปข้างหน้า" OR "ปุ่มClear",
                           PV := 1);
   IF "IEC_Counter_0_DB_672".Q THEN #Output := 198; END_IF;
   "IEC_Counter_0_DB_671".CTU(CU := ("ยา 199" = 1) AND ("IEC_Counter_0_DB_671".CV < 1),
                           R := "Stepper Motor ทำงาน สั่งconveyor เคลื่อที่ไปข้างหน้า" OR "ปุ่มClear",
                           PV := 1);
   IF "IEC_Counter_0_DB_671".Q THEN #Output := 199; END_IF;
   "IEC_Counter_0_DB_670".CTU(CU := ("ยา 200" = 1) AND ("IEC_Counter_0_DB_670".CV < 1),
                           R := "Stepper Motor ทำงาน สั่งconveyor เคลื่อที่ไปข้างหน้า" OR "ปุ่มClear",
                           PV := 1);
   IF "IEC_Counter_0_DB_670".Q THEN #Output := 200; END_IF;
END_REGION

REGION Network 11
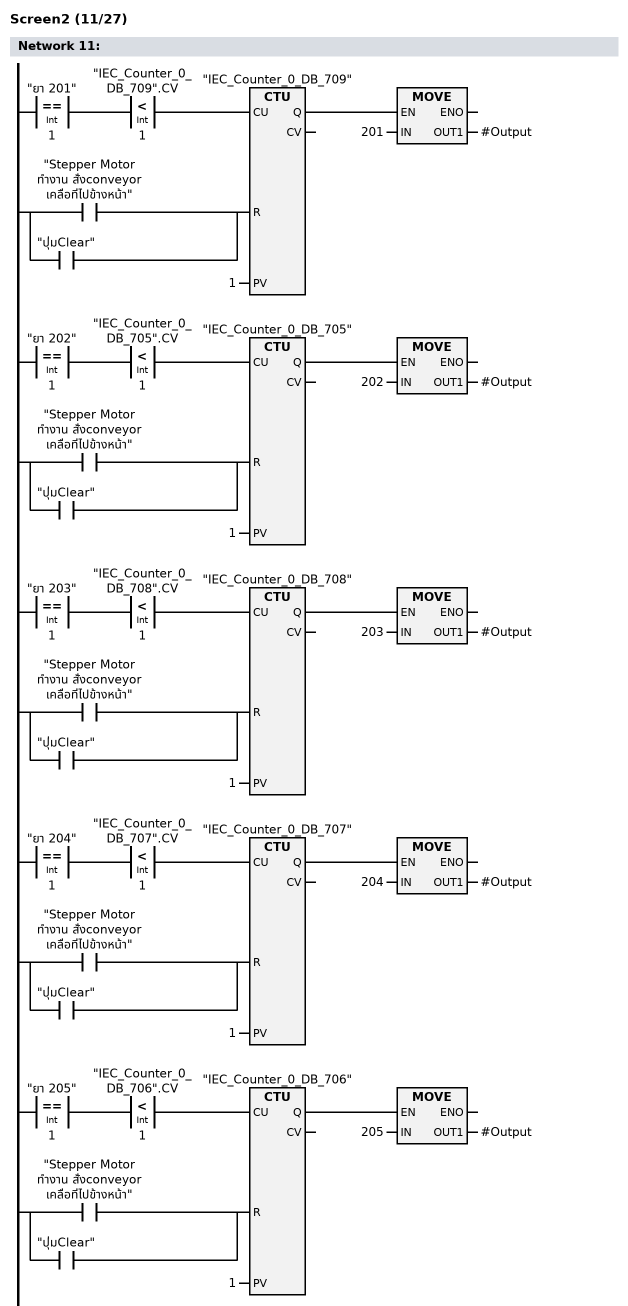
